{region "07 - Consume Start and Abort without restarting"}
FSteps[7].ExpectedState := E_State.Completed;
FSteps[7].ExpectedResult := E_Result.Passed;
FSteps[7].ExpectedReady := FALSE;
FSteps[7].ExpectedPassedCount := 2;
FSteps[7].ExpectedFailedCount := 0;
FSteps[7].CheckFinalization := TRUE;
FSteps[7].ExpectedFinalizationCount := 1;
FSteps[7].ExpectedCompletionCount := 1;
FSteps[7].ExpectedFinalResult := E_Result.Passed;
FSteps[7].ExpectRuntimeHeld := TRUE;
FSteps[7].RequestStart := TRUE;
FSteps[7].RequestAbort := TRUE;
FSteps[7].ExpectedHookCount := 1;
FSteps[7].ExpectedHooks[1].Hook := E_LifecycleHook.Aggregate;
FSteps[7].ExpectedHooks[1].State := E_State.Completed;
FSteps[7].ExpectedHooks[1].Enabled := TRUE;
{endregion}

{region "08 - Remain quiet after rejected terminal requests"}
FSteps[8].ExpectedState := E_State.Completed;
FSteps[8].ExpectedResult := E_Result.Passed;
FSteps[8].ExpectedReady := FALSE;
FSteps[8].ExpectedPassedCount := 2;
FSteps[8].ExpectedFailedCount := 0;
FSteps[8].CheckFinalization := TRUE;
FSteps[8].ExpectedFinalizationCount := 1;
FSteps[8].ExpectedCompletionCount := 1;
FSteps[8].ExpectedFinalResult := E_Result.Passed;
FSteps[8].ExpectRuntimeHeld := TRUE;
FSteps[8].ExpectQuietCall := TRUE;
FSteps[8].ExpectedHookCount := 1;
FSteps[8].ExpectedHooks[1].Hook := E_LifecycleHook.Aggregate;
FSteps[8].ExpectedHooks[1].State := E_State.Completed;
FSteps[8].ExpectedHooks[1].Enabled := TRUE;
{endregion}

{region "09 - Reset clears the first result and competing requests"}
FSteps[9].ExpectedState := E_State.Idle;
FSteps[9].ExpectedResult := E_Result.NotEvaluated;
FSteps[9].ExpectedReady := TRUE;
FSteps[9].ExpectedPassedCount := 0;
FSteps[9].ExpectedFailedCount := 0;
FSteps[9].CheckFinalization := TRUE;
FSteps[9].ExpectedFinalizationCount := 1;
FSteps[9].ExpectedCompletionCount := 1;
FSteps[9].ExpectedFinalResult := E_Result.Passed;
FSteps[9].RequestReset := TRUE;
FSteps[9].RequestStart := TRUE;
FSteps[9].RequestAbort := TRUE;
FSteps[9].ExpectRuntimeCleared := TRUE;
FSteps[9].ExpectedHookCount := 6;
FSteps[9].ExpectedHooks[1].Hook := E_LifecycleHook.Reset;
FSteps[9].ExpectedHooks[1].State := E_State.Reset;
FSteps[9].ExpectedHooks[1].Enabled := TRUE;
FSteps[9].ExpectedHooks[2].Hook := E_LifecycleHook.Abort;
FSteps[9].ExpectedHooks[2].State := E_State.Idle;
FSteps[9].ExpectedHooks[2].Enabled := FALSE;
FSteps[9].ExpectedHooks[3].Hook := E_LifecycleHook.Preparations;
FSteps[9].ExpectedHooks[3].State := E_State.Idle;
FSteps[9].ExpectedHooks[3].Enabled := FALSE;
FSteps[9].ExpectedHooks[4].Hook := E_LifecycleHook.Tests;
FSteps[9].ExpectedHooks[4].State := E_State.Idle;
FSteps[9].ExpectedHooks[4].Enabled := FALSE;
FSteps[9].ExpectedHooks[5].Hook := E_LifecycleHook.Assertions;
FSteps[9].ExpectedHooks[5].State := E_State.Idle;
FSteps[9].ExpectedHooks[5].Enabled := FALSE;
FSteps[9].ExpectedHooks[6].Hook := E_LifecycleHook.Aggregate;
FSteps[9].ExpectedHooks[6].State := E_State.Idle;
FSteps[9].ExpectedHooks[6].Enabled := TRUE;
{endregion}

{region "10 - Do not retain a Start from the Reset call"}
FSteps[10].ExpectedState := E_State.Idle;
FSteps[10].ExpectedResult := E_Result.NotEvaluated;
FSteps[10].ExpectedReady := TRUE;
FSteps[10].ExpectedPassedCount := 0;
FSteps[10].ExpectedFailedCount := 0;
FSteps[10].CheckFinalization := TRUE;
FSteps[10].ExpectedFinalizationCount := 1;
FSteps[10].ExpectedCompletionCount := 1;
FSteps[10].ExpectedFinalResult := E_Result.Passed;
FSteps[10].ExpectRuntimeCleared := TRUE;
FSteps[10].ExpectQuietCall := TRUE;
FSteps[10].ExpectedHookCount := 5;
FSteps[10].ExpectedHooks[1].Hook := E_LifecycleHook.Abort;
FSteps[10].ExpectedHooks[1].State := E_State.Idle;
FSteps[10].ExpectedHooks[1].Enabled := FALSE;
FSteps[10].ExpectedHooks[2].Hook := E_LifecycleHook.Preparations;
FSteps[10].ExpectedHooks[2].State := E_State.Idle;
FSteps[10].ExpectedHooks[2].Enabled := FALSE;
FSteps[10].ExpectedHooks[3].Hook := E_LifecycleHook.Tests;
FSteps[10].ExpectedHooks[3].State := E_State.Idle;
FSteps[10].ExpectedHooks[3].Enabled := FALSE;
FSteps[10].ExpectedHooks[4].Hook := E_LifecycleHook.Assertions;
FSteps[10].ExpectedHooks[4].State := E_State.Idle;
FSteps[10].ExpectedHooks[4].Enabled := FALSE;
FSteps[10].ExpectedHooks[5].Hook := E_LifecycleHook.Aggregate;
FSteps[10].ExpectedHooks[5].State := E_State.Idle;
FSteps[10].ExpectedHooks[5].Enabled := TRUE;
{endregion}

{region "11 - Start a fresh second execution"}
FSteps[11].ExpectedState := E_State.Starting;
FSteps[11].ExpectedResult := E_Result.NotEvaluated;
FSteps[11].ExpectedReady := FALSE;
FSteps[11].ExpectedPassedCount := 0;
FSteps[11].ExpectedFailedCount := 0;
FSteps[11].CheckFinalization := TRUE;
FSteps[11].ExpectedFinalizationCount := 1;
FSteps[11].ExpectedCompletionCount := 1;
FSteps[11].ExpectedFinalResult := E_Result.Passed;
FSteps[11].RequestStart := TRUE;
FSteps[11].ExpectedHookCount := 5;
FSteps[11].ExpectedHooks[1].Hook := E_LifecycleHook.Abort;
FSteps[11].ExpectedHooks[1].State := E_State.Starting;
FSteps[11].ExpectedHooks[1].Enabled := FALSE;
FSteps[11].ExpectedHooks[2].Hook := E_LifecycleHook.Preparations;
FSteps[11].ExpectedHooks[2].State := E_State.Starting;
FSteps[11].ExpectedHooks[2].Enabled := FALSE;
FSteps[11].ExpectedHooks[3].Hook := E_LifecycleHook.Tests;
FSteps[11].ExpectedHooks[3].State := E_State.Starting;
FSteps[11].ExpectedHooks[3].Enabled := FALSE;
FSteps[11].ExpectedHooks[4].Hook := E_LifecycleHook.Assertions;
FSteps[11].ExpectedHooks[4].State := E_State.Starting;
FSteps[11].ExpectedHooks[4].Enabled := FALSE;
FSteps[11].ExpectedHooks[5].Hook := E_LifecycleHook.Aggregate;
FSteps[11].ExpectedHooks[5].State := E_State.Starting;
FSteps[11].ExpectedHooks[5].Enabled := TRUE;
{endregion}

{region "12 - Both Assertions pass after Reset"}
FSteps[12].ExpectedState := E_State.Running;
FSteps[12].ExpectedResult := E_Result.NotEvaluated;
FSteps[12].ExpectedReady := FALSE;
FSteps[12].ExpectedPassedCount := 2;
FSteps[12].ExpectedFailedCount := 0;
FSteps[12].CheckFinalization := TRUE;
FSteps[12].ExpectedFinalizationCount := 1;
FSteps[12].ExpectedCompletionCount := 1;
FSteps[12].ExpectedFinalResult := E_Result.Passed;
FSteps[12].ExpectedHookCount := 5;
FSteps[12].ExpectedHooks[1].Hook := E_LifecycleHook.Abort;
FSteps[12].ExpectedHooks[1].State := E_State.Running;
FSteps[12].ExpectedHooks[1].Enabled := FALSE;
FSteps[12].ExpectedHooks[2].Hook := E_LifecycleHook.Preparations;
FSteps[12].ExpectedHooks[2].State := E_State.Running;
FSteps[12].ExpectedHooks[2].Enabled := FALSE;
FSteps[12].ExpectedHooks[3].Hook := E_LifecycleHook.Tests;
FSteps[12].ExpectedHooks[3].State := E_State.Running;
FSteps[12].ExpectedHooks[3].Enabled := TRUE;
FSteps[12].ExpectedHooks[4].Hook := E_LifecycleHook.Assertions;
FSteps[12].ExpectedHooks[4].State := E_State.Running;
FSteps[12].ExpectedHooks[4].Enabled := TRUE;
FSteps[12].ExpectedHooks[5].Hook := E_LifecycleHook.Aggregate;
FSteps[12].ExpectedHooks[5].State := E_State.Running;
FSteps[12].ExpectedHooks[5].Enabled := TRUE;
{endregion}

{region "13 - Publish a new successful finalization"}
FSteps[13].ExpectedState := E_State.Completing;
FSteps[13].ExpectedResult := E_Result.Passed;
FSteps[13].ExpectedReady := FALSE;
FSteps[13].ExpectedPassedCount := 2;
FSteps[13].ExpectedFailedCount := 0;
FSteps[13].FinishTests := TRUE;
FSteps[13].CheckFinalization := TRUE;
FSteps[13].ExpectedFinalizationCount := 2;
FSteps[13].ExpectedCompletionCount := 1;
FSteps[13].ExpectedFinalResult := E_Result.Passed;
FSteps[13].ExpectedHookCount := 5;
FSteps[13].ExpectedHooks[1].Hook := E_LifecycleHook.Abort;
FSteps[13].ExpectedHooks[1].State := E_State.Running;
FSteps[13].ExpectedHooks[1].Enabled := FALSE;
FSteps[13].ExpectedHooks[2].Hook := E_LifecycleHook.Preparations;
FSteps[13].ExpectedHooks[2].State := E_State.Running;
FSteps[13].ExpectedHooks[2].Enabled := FALSE;
FSteps[13].ExpectedHooks[3].Hook := E_LifecycleHook.Tests;
FSteps[13].ExpectedHooks[3].State := E_State.Running;
FSteps[13].ExpectedHooks[3].Enabled := TRUE;
FSteps[13].ExpectedHooks[4].Hook := E_LifecycleHook.Assertions;
FSteps[13].ExpectedHooks[4].State := E_State.Completing;
FSteps[13].ExpectedHooks[4].Enabled := FALSE;
FSteps[13].ExpectedHooks[5].Hook := E_LifecycleHook.Aggregate;
FSteps[13].ExpectedHooks[5].State := E_State.Completing;
FSteps[13].ExpectedHooks[5].Enabled := TRUE;
{endregion}

{region "14 - Complete the second execution"}
FSteps[14].ExpectedState := E_State.Completed;
FSteps[14].ExpectedResult := E_Result.Passed;
FSteps[14].ExpectedReady := FALSE;
FSteps[14].ExpectedPassedCount := 2;
FSteps[14].ExpectedFailedCount := 0;
FSteps[14].ExpectRuntimeHeld := TRUE;
FSteps[14].CheckFinalization := TRUE;
FSteps[14].ExpectedFinalizationCount := 2;
FSteps[14].ExpectedCompletionCount := 2;
FSteps[14].ExpectedFinalResult := E_Result.Passed;
FSteps[14].ExpectedHookCount := 1;
FSteps[14].ExpectedHooks[1].Hook := E_LifecycleHook.Aggregate;
FSteps[14].ExpectedHooks[1].State := E_State.Completed;
FSteps[14].ExpectedHooks[1].Enabled := TRUE;
{endregion}

{region "15 - Do not repeat second-run finalization"}
FSteps[15].ExpectedState := E_State.Completed;
FSteps[15].ExpectedResult := E_Result.Passed;
FSteps[15].ExpectedReady := FALSE;
FSteps[15].ExpectedPassedCount := 2;
FSteps[15].ExpectedFailedCount := 0;
FSteps[15].ExpectQuietCall := TRUE;
FSteps[15].ExpectRuntimeHeld := TRUE;
FSteps[15].CheckFinalization := TRUE;
FSteps[15].ExpectedFinalizationCount := 2;
FSteps[15].ExpectedCompletionCount := 2;
FSteps[15].ExpectedFinalResult := E_Result.Passed;
FSteps[15].ExpectedHookCount := 1;
FSteps[15].ExpectedHooks[1].Hook := E_LifecycleHook.Aggregate;
FSteps[15].ExpectedHooks[1].State := E_State.Completed;
FSteps[15].ExpectedHooks[1].Enabled := TRUE;
{endregion}
END_METHOD

END_FUNCTION_BLOCK

// ---- SelfTests/TestCases/TestSuite_TestCaseLifecycle/Test_LifecycleRepeatAfterFailed.TcPOU
{region 'Documentation'}
(*!
<summary>Checks stable Failed completion, one-shot finalization and a fresh successful run after Reset.</summary>
*)
{endregion}
FUNCTION_BLOCK Test_LifecycleRepeatAfterFailed EXTENDS TestCaseLifecycleTestBase

SUPER^();

{region 'Documentation'}
(*!
<summary>Defines two independent run outcomes and cumulative event expectations across Reset.</summary>
*)
{endregion}
METHOD PROTECTED ConfigureScenario
FSubjectPreparationCount := 0;
FSubjectTestCount := 1;
FStepCount := 15;

{region "01 - Reset establishes the initial Idle state"}
FSteps[1].ExpectedState := E_State.Idle;
FSteps[1].ExpectedResult := E_Result.NotEvaluated;
FSteps[1].ExpectedReady := TRUE;
FSteps[1].ExpectedPassedCount := 0;
FSteps[1].ExpectedFailedCount := 0;
FSteps[1].RequestReset := TRUE;
FSteps[1].ExpectRuntimeCleared := TRUE;
FSteps[1].CheckFinalization := TRUE;
FSteps[1].ExpectedFinalizationCount := 0;
FSteps[1].ExpectedCompletionCount := 0;
FSteps[1].ExpectedFinalResult := E_Result.Failed;
FSteps[1].ExpectedHookCount := 6;
FSteps[1].ExpectedHooks[1].Hook := E_LifecycleHook.Reset;
FSteps[1].ExpectedHooks[1].State := E_State.Reset;
FSteps[1].ExpectedHooks[1].Enabled := TRUE;
FSteps[1].ExpectedHooks[2].Hook := E_LifecycleHook.Abort;
FSteps[1].ExpectedHooks[2].State := E_State.Idle;
FSteps[1].ExpectedHooks[2].Enabled := FALSE;
FSteps[1].ExpectedHooks[3].Hook := E_LifecycleHook.Preparations;
FSteps[1].ExpectedHooks[3].State := E_State.Idle;
FSteps[1].ExpectedHooks[3].Enabled := FALSE;
FSteps[1].ExpectedHooks[4].Hook := E_LifecycleHook.Tests;
FSteps[1].ExpectedHooks[4].State := E_State.Idle;
FSteps[1].ExpectedHooks[4].Enabled := FALSE;
FSteps[1].ExpectedHooks[5].Hook := E_LifecycleHook.Assertions;
FSteps[1].ExpectedHooks[5].State := E_State.Idle;
FSteps[1].ExpectedHooks[5].Enabled := FALSE;
FSteps[1].ExpectedHooks[6].Hook := E_LifecycleHook.Aggregate;
FSteps[1].ExpectedHooks[6].State := E_State.Idle;
FSteps[1].ExpectedHooks[6].Enabled := TRUE;
{endregion}

{region "02 - Start the first execution"}
FSteps[2].ExpectedState := E_State.Starting;
FSteps[2].ExpectedResult := E_Result.NotEvaluated;
FSteps[2].ExpectedReady := FALSE;
FSteps[2].ExpectedPassedCount := 0;
FSteps[2].ExpectedFailedCount := 0;
FSteps[2].RequestStart := TRUE;
FSteps[2].CheckFinalization := TRUE;
FSteps[2].ExpectedFinalizationCount := 0;
FSteps[2].ExpectedCompletionCount := 0;
FSteps[2].ExpectedFinalResult := E_Result.Failed;
FSteps[2].ExpectedHookCount := 5;
FSteps[2].ExpectedHooks[1].Hook := E_LifecycleHook.Abort;
FSteps[2].ExpectedHooks[1].State := E_State.Starting;
FSteps[2].ExpectedHooks[1].Enabled := FALSE;
FSteps[2].ExpectedHooks[2].Hook := E_LifecycleHook.Preparations;
FSteps[2].ExpectedHooks[2].State := E_State.Starting;
FSteps[2].ExpectedHooks[2].Enabled := FALSE;
FSteps[2].ExpectedHooks[3].Hook := E_LifecycleHook.Tests;
FSteps[2].ExpectedHooks[3].State := E_State.Starting;
FSteps[2].ExpectedHooks[3].Enabled := FALSE;
FSteps[2].ExpectedHooks[4].Hook := E_LifecycleHook.Assertions;
FSteps[2].ExpectedHooks[4].State := E_State.Starting;
FSteps[2].ExpectedHooks[4].Enabled := FALSE;
FSteps[2].ExpectedHooks[5].Hook := E_LifecycleHook.Aggregate;
FSteps[2].ExpectedHooks[5].State := E_State.Starting;
FSteps[2].ExpectedHooks[5].Enabled := TRUE;
{endregion}

{region "03 - Evaluate both child Assertions"}
FSteps[3].ExpectedState := E_State.Running;
FSteps[3].ExpectedResult := E_Result.NotEvaluated;
FSteps[3].ExpectedReady := FALSE;
FSteps[3].ExpectedPassedCount := 1;
FSteps[3].ExpectedFailedCount := 1;
FSteps[3].AssertionCondition := FALSE;
FSteps[3].CheckFinalization := TRUE;
FSteps[3].ExpectedFinalizationCount := 0;
FSteps[3].ExpectedCompletionCount := 0;
FSteps[3].ExpectedFinalResult := E_Result.Failed;
FSteps[3].ExpectedHookCount := 5;
FSteps[3].ExpectedHooks[1].Hook := E_LifecycleHook.Abort;
FSteps[3].ExpectedHooks[1].State := E_State.Running;
FSteps[3].ExpectedHooks[1].Enabled := FALSE;
FSteps[3].ExpectedHooks[2].Hook := E_LifecycleHook.Preparations;
FSteps[3].ExpectedHooks[2].State := E_State.Running;
FSteps[3].ExpectedHooks[2].Enabled := FALSE;
FSteps[3].ExpectedHooks[3].Hook := E_LifecycleHook.Tests;
FSteps[3].ExpectedHooks[3].State := E_State.Running;
FSteps[3].ExpectedHooks[3].Enabled := TRUE;
FSteps[3].ExpectedHooks[4].Hook := E_LifecycleHook.Assertions;
FSteps[3].ExpectedHooks[4].State := E_State.Running;
FSteps[3].ExpectedHooks[4].Enabled := TRUE;
FSteps[3].ExpectedHooks[5].Hook := E_LifecycleHook.Aggregate;
FSteps[3].ExpectedHooks[5].State := E_State.Running;
FSteps[3].ExpectedHooks[5].Enabled := TRUE;
{endregion}

{region "04 - Finalize the first result"}
FSteps[4].ExpectedState := E_State.Completing;
FSteps[4].ExpectedResult := E_Result.Failed;
FSteps[4].ExpectedReady := FALSE;
FSteps[4].ExpectedPassedCount := 1;
FSteps[4].ExpectedFailedCount := 1;
FSteps[4].FinishTests := TRUE;
FSteps[4].CheckFinalization := TRUE;
FSteps[4].ExpectedFinalizationCount := 1;
FSteps[4].ExpectedCompletionCount := 0;
FSteps[4].ExpectedFinalResult := E_Result.Failed;
FSteps[4].ExpectedHookCount := 5;
FSteps[4].ExpectedHooks[1].Hook := E_LifecycleHook.Abort;
FSteps[4].ExpectedHooks[1].State := E_State.Running;
FSteps[4].ExpectedHooks[1].Enabled := FALSE;
FSteps[4].ExpectedHooks[2].Hook := E_LifecycleHook.Preparations;
FSteps[4].ExpectedHooks[2].State := E_State.Running;
FSteps[4].ExpectedHooks[2].Enabled := FALSE;
FSteps[4].ExpectedHooks[3].Hook := E_LifecycleHook.Tests;
FSteps[4].ExpectedHooks[3].State := E_State.Running;
FSteps[4].ExpectedHooks[3].Enabled := TRUE;
FSteps[4].ExpectedHooks[4].Hook := E_LifecycleHook.Assertions;
FSteps[4].ExpectedHooks[4].State := E_State.Completing;
FSteps[4].ExpectedHooks[4].Enabled := FALSE;
FSteps[4].ExpectedHooks[5].Hook := E_LifecycleHook.Aggregate;
FSteps[4].ExpectedHooks[5].State := E_State.Completing;
FSteps[4].ExpectedHooks[5].Enabled := TRUE;
{endregion}

{region "05 - Observe the final Completed transition"}
FSteps[5].ExpectedState := E_State.Completed;
FSteps[5].ExpectedResult := E_Result.Failed;
FSteps[5].ExpectedReady := FALSE;
FSteps[5].ExpectedPassedCount := 1;
FSteps[5].ExpectedFailedCount := 1;
FSteps[5].CheckFinalization := TRUE;
FSteps[5].ExpectedFinalizationCount := 1;
FSteps[5].ExpectedCompletionCount := 1;
FSteps[5].ExpectedFinalResult := E_Result.Failed;
FSteps[5].ExpectRuntimeHeld := TRUE;
FSteps[5].ExpectedHookCount := 1;
FSteps[5].ExpectedHooks[1].Hook := E_LifecycleHook.Aggregate;
FSteps[5].ExpectedHooks[1].State := E_State.Completed;
FSteps[5].ExpectedHooks[1].Enabled := TRUE;
{endregion}

{region "06 - Ignore processing inputs while Completed"}
FSteps[6].ExpectedState := E_State.Completed;
FSteps[6].ExpectedResult := E_Result.Failed;
FSteps[6].ExpectedReady := FALSE;
FSteps[6].ExpectedPassedCount := 1;
FSteps[6].ExpectedFailedCount := 1;
FSteps[6].CheckFinalization := TRUE;
FSteps[6].ExpectedFinalizationCount := 1;
FSteps[6].ExpectedCompletionCount := 1;
FSteps[6].ExpectedFinalResult := E_Result.Failed;
FSteps[6].ExpectRuntimeHeld := TRUE;
FSteps[6].ExpectQuietCall := TRUE;
FSteps[6].Ready := FALSE;
FSteps[6].ResetError := TRUE;
FSteps[6].AbortError := TRUE;
FSteps[6].TestError := TRUE;
FSteps[6].PreparationError := TRUE;
FSteps[6].AdvancePreparation := TRUE;
FSteps[6].FinishPreparations := TRUE;
FSteps[6].AdvanceTest := TRUE;
FSteps[6].FinishTests := TRUE;
FSteps[6].AssertionCondition := FALSE;
FSteps[6].ExpectedHookCount := 1;
FSteps[6].ExpectedHooks[1].Hook := E_LifecycleHook.Aggregate;
FSteps[6].ExpectedHooks[1].State := E_State.Completed;
FSteps[6].ExpectedHooks[1].Enabled := TRUE;
{endregion}

{region "07 - Consume Start and Abort without restarting"}
FSteps[7].ExpectedState := E_State.Completed;
FSteps[7].ExpectedResult := E_Result.Failed;
FSteps[7].ExpectedReady := FALSE;
FSteps[7].ExpectedPassedCount := 1;
FSteps[7].ExpectedFailedCount := 1;
FSteps[7].CheckFinalization := TRUE;
FSteps[7].ExpectedFinalizationCount := 1;
FSteps[7].ExpectedCompletionCount := 1;
FSteps[7].ExpectedFinalResult := E_Result.Failed;
FSteps[7].ExpectRuntimeHeld := TRUE;
FSteps[7].RequestStart := TRUE;
FSteps[7].RequestAbort := TRUE;
FSteps[7].ExpectedHookCount := 1;
FSteps[7].ExpectedHooks[1].Hook := E_LifecycleHook.Aggregate;
FSteps[7].ExpectedHooks[1].State := E_State.Completed;
FSteps[7].ExpectedHooks[1].Enabled := TRUE;
{endregion}

{region "08 - Remain quiet after rejected terminal requests"}
FSteps[8].ExpectedState := E_State.Completed;
FSteps[8].ExpectedResult := E_Result.Failed;
FSteps[8].ExpectedReady := FALSE;
FSteps[8].ExpectedPassedCount := 1;
FSteps[8].ExpectedFailedCount := 1;
FSteps[8].CheckFinalization := TRUE;
FSteps[8].ExpectedFinalizationCount := 1;
FSteps[8].ExpectedCompletionCount := 1;
FSteps[8].ExpectedFinalResult := E_Result.Failed;
FSteps[8].ExpectRuntimeHeld := TRUE;
FSteps[8].ExpectQuietCall := TRUE;
FSteps[8].ExpectedHookCount := 1;
FSteps[8].ExpectedHooks[1].Hook := E_LifecycleHook.Aggregate;
FSteps[8].ExpectedHooks[1].State := E_State.Completed;
FSteps[8].ExpectedHooks[1].Enabled := TRUE;
{endregion}

{region "09 - Reset clears the first result and competing requests"}
FSteps[9].ExpectedState := E_State.Idle;
FSteps[9].ExpectedResult := E_Result.NotEvaluated;
FSteps[9].ExpectedReady := TRUE;
FSteps[9].ExpectedPassedCount := 0;
FSteps[9].ExpectedFailedCount := 0;
FSteps[9].CheckFinalization := TRUE;
FSteps[9].ExpectedFinalizationCount := 1;
FSteps[9].ExpectedCompletionCount := 1;
FSteps[9].ExpectedFinalResult := E_Result.Failed;
FSteps[9].RequestReset := TRUE;
FSteps[9].RequestStart := TRUE;
FSteps[9].RequestAbort := TRUE;
FSteps[9].ExpectRuntimeCleared := TRUE;
FSteps[9].ExpectedHookCount := 6;
FSteps[9].ExpectedHooks[1].Hook := E_LifecycleHook.Reset;
FSteps[9].ExpectedHooks[1].State := E_State.Reset;
FSteps[9].ExpectedHooks[1].Enabled := TRUE;
FSteps[9].ExpectedHooks[2].Hook := E_LifecycleHook.Abort;
FSteps[9].ExpectedHooks[2].State := E_State.Idle;
FSteps[9].ExpectedHooks[2].Enabled := FALSE;
FSteps[9].ExpectedHooks[3].Hook := E_LifecycleHook.Preparations;
FSteps[9].ExpectedHooks[3].State := E_State.Idle;
FSteps[9].ExpectedHooks[3].Enabled := FALSE;
FSteps[9].ExpectedHooks[4].Hook := E_LifecycleHook.Tests;
FSteps[9].ExpectedHooks[4].State := E_State.Idle;
FSteps[9].ExpectedHooks[4].Enabled := FALSE;
FSteps[9].ExpectedHooks[5].Hook := E_LifecycleHook.Assertions;
FSteps[9].ExpectedHooks[5].State := E_State.Idle;
FSteps[9].ExpectedHooks[5].Enabled := FALSE;
FSteps[9].ExpectedHooks[6].Hook := E_LifecycleHook.Aggregate;
FSteps[9].ExpectedHooks[6].State := E_State.Idle;
FSteps[9].ExpectedHooks[6].Enabled := TRUE;
{endregion}

{region "10 - Do not retain a Start from the Reset call"}
FSteps[10].ExpectedState := E_State.Idle;
FSteps[10].ExpectedResult := E_Result.NotEvaluated;
FSteps[10].ExpectedReady := TRUE;
FSteps[10].ExpectedPassedCount := 0;
FSteps[10].ExpectedFailedCount := 0;
FSteps[10].CheckFinalization := TRUE;
FSteps[10].ExpectedFinalizationCount := 1;
FSteps[10].ExpectedCompletionCount := 1;
FSteps[10].ExpectedFinalResult := E_Result.Failed;
FSteps[10].ExpectRuntimeCleared := TRUE;
FSteps[10].ExpectQuietCall := TRUE;
FSteps[10].ExpectedHookCount := 5;
FSteps[10].ExpectedHooks[1].Hook := E_LifecycleHook.Abort;
FSteps[10].ExpectedHooks[1].State := E_State.Idle;
FSteps[10].ExpectedHooks[1].Enabled := FALSE;
FSteps[10].ExpectedHooks[2].Hook := E_LifecycleHook.Preparations;
FSteps[10].ExpectedHooks[2].State := E_State.Idle;
FSteps[10].ExpectedHooks[2].Enabled := FALSE;
FSteps[10].ExpectedHooks[3].Hook := E_LifecycleHook.Tests;
FSteps[10].ExpectedHooks[3].State := E_State.Idle;
FSteps[10].ExpectedHooks[3].Enabled := FALSE;
FSteps[10].ExpectedHooks[4].Hook := E_LifecycleHook.Assertions;
FSteps[10].ExpectedHooks[4].State := E_State.Idle;
FSteps[10].ExpectedHooks[4].Enabled := FALSE;
FSteps[10].ExpectedHooks[5].Hook := E_LifecycleHook.Aggregate;
FSteps[10].ExpectedHooks[5].State := E_State.Idle;
FSteps[10].ExpectedHooks[5].Enabled := TRUE;
{endregion}

{region "11 - Start a fresh second execution"}
FSteps[11].ExpectedState := E_State.Starting;
FSteps[11].ExpectedResult := E_Result.NotEvaluated;
FSteps[11].ExpectedReady := FALSE;
FSteps[11].ExpectedPassedCount := 0;
FSteps[11].ExpectedFailedCount := 0;
FSteps[11].CheckFinalization := TRUE;
FSteps[11].ExpectedFinalizationCount := 1;
FSteps[11].ExpectedCompletionCount := 1;
FSteps[11].ExpectedFinalResult := E_Result.Failed;
FSteps[11].RequestStart := TRUE;
FSteps[11].ExpectedHookCount := 5;
FSteps[11].ExpectedHooks[1].Hook := E_LifecycleHook.Abort;
FSteps[11].ExpectedHooks[1].State := E_State.Starting;
FSteps[11].ExpectedHooks[1].Enabled := FALSE;
FSteps[11].ExpectedHooks[2].Hook := E_LifecycleHook.Preparations;
FSteps[11].ExpectedHooks[2].State := E_State.Starting;
FSteps[11].ExpectedHooks[2].Enabled := FALSE;
FSteps[11].ExpectedHooks[3].Hook := E_LifecycleHook.Tests;
FSteps[11].ExpectedHooks[3].State := E_State.Starting;
FSteps[11].ExpectedHooks[3].Enabled := FALSE;
FSteps[11].ExpectedHooks[4].Hook := E_LifecycleHook.Assertions;
FSteps[11].ExpectedHooks[4].State := E_State.Starting;
FSteps[11].ExpectedHooks[4].Enabled := FALSE;
FSteps[11].ExpectedHooks[5].Hook := E_LifecycleHook.Aggregate;
FSteps[11].ExpectedHooks[5].State := E_State.Starting;
FSteps[11].ExpectedHooks[5].Enabled := TRUE;
{endregion}

{region "12 - Both Assertions pass after Reset"}
FSteps[12].ExpectedState := E_State.Running;
FSteps[12].ExpectedResult := E_Result.NotEvaluated;
FSteps[12].ExpectedReady := FALSE;
FSteps[12].ExpectedPassedCount := 2;
FSteps[12].ExpectedFailedCount := 0;
FSteps[12].CheckFinalization := TRUE;
FSteps[12].ExpectedFinalizationCount := 1;
FSteps[12].ExpectedCompletionCount := 1;
FSteps[12].ExpectedFinalResult := E_Result.Failed;
FSteps[12].ExpectedHookCount := 5;
FSteps[12].ExpectedHooks[1].Hook := E_LifecycleHook.Abort;
FSteps[12].ExpectedHooks[1].State := E_State.Running;
FSteps[12].ExpectedHooks[1].Enabled := FALSE;
FSteps[12].ExpectedHooks[2].Hook := E_LifecycleHook.Preparations;
FSteps[12].ExpectedHooks[2].State := E_State.Running;
FSteps[12].ExpectedHooks[2].Enabled := FALSE;
FSteps[12].ExpectedHooks[3].Hook := E_LifecycleHook.Tests;
FSteps[12].ExpectedHooks[3].State := E_State.Running;
FSteps[12].ExpectedHooks[3].Enabled := TRUE;
FSteps[12].ExpectedHooks[4].Hook := E_LifecycleHook.Assertions;
FSteps[12].ExpectedHooks[4].State := E_State.Running;
FSteps[12].ExpectedHooks[4].Enabled := TRUE;
FSteps[12].ExpectedHooks[5].Hook := E_LifecycleHook.Aggregate;
FSteps[12].ExpectedHooks[5].State := E_State.Running;
FSteps[12].ExpectedHooks[5].Enabled := TRUE;
{endregion}

{region "13 - Publish a new successful finalization"}
FSteps[13].ExpectedState := E_State.Completing;
FSteps[13].ExpectedResult := E_Result.Passed;
FSteps[13].ExpectedReady := FALSE;
FSteps[13].ExpectedPassedCount := 2;
FSteps[13].ExpectedFailedCount := 0;
FSteps[13].FinishTests := TRUE;
FSteps[13].CheckFinalization := TRUE;
FSteps[13].ExpectedFinalizationCount := 2;
FSteps[13].ExpectedCompletionCount := 1;
FSteps[13].ExpectedFinalResult := E_Result.Passed;
FSteps[13].ExpectedHookCount := 5;
FSteps[13].ExpectedHooks[1].Hook := E_LifecycleHook.Abort;
FSteps[13].ExpectedHooks[1].State := E_State.Running;
FSteps[13].ExpectedHooks[1].Enabled := FALSE;
FSteps[13].ExpectedHooks[2].Hook := E_LifecycleHook.Preparations;
FSteps[13].ExpectedHooks[2].State := E_State.Running;
FSteps[13].ExpectedHooks[2].Enabled := FALSE;
FSteps[13].ExpectedHooks[3].Hook := E_LifecycleHook.Tests;
FSteps[13].ExpectedHooks[3].State := E_State.Running;
FSteps[13].ExpectedHooks[3].Enabled := TRUE;
FSteps[13].ExpectedHooks[4].Hook := E_LifecycleHook.Assertions;
FSteps[13].ExpectedHooks[4].State := E_State.Completing;
FSteps[13].ExpectedHooks[4].Enabled := FALSE;
FSteps[13].ExpectedHooks[5].Hook := E_LifecycleHook.Aggregate;
FSteps[13].ExpectedHooks[5].State := E_State.Completing;
FSteps[13].ExpectedHooks[5].Enabled := TRUE;
{endregion}

{region "14 - Complete the second execution"}
FSteps[14].ExpectedState := E_State.Completed;
FSteps[14].ExpectedResult := E_Result.Passed;
FSteps[14].ExpectedReady := FALSE;
FSteps[14].ExpectedPassedCount := 2;
FSteps[14].ExpectedFailedCount := 0;
FSteps[14].ExpectRuntimeHeld := TRUE;
FSteps[14].CheckFinalization := TRUE;
FSteps[14].ExpectedFinalizationCount := 2;
FSteps[14].ExpectedCompletionCount := 2;
FSteps[14].ExpectedFinalResult := E_Result.Passed;
FSteps[14].ExpectedHookCount := 1;
FSteps[14].ExpectedHooks[1].Hook := E_LifecycleHook.Aggregate;
FSteps[14].ExpectedHooks[1].State := E_State.Completed;
FSteps[14].ExpectedHooks[1].Enabled := TRUE;
{endregion}

{region "15 - Do not repeat second-run finalization"}
FSteps[15].ExpectedState := E_State.Completed;
FSteps[15].ExpectedResult := E_Result.Passed;
FSteps[15].ExpectedReady := FALSE;
FSteps[15].ExpectedPassedCount := 2;
FSteps[15].ExpectedFailedCount := 0;
FSteps[15].ExpectQuietCall := TRUE;
FSteps[15].ExpectRuntimeHeld := TRUE;
FSteps[15].CheckFinalization := TRUE;
FSteps[15].ExpectedFinalizationCount := 2;
FSteps[15].ExpectedCompletionCount := 2;
FSteps[15].ExpectedFinalResult := E_Result.Passed;
FSteps[15].ExpectedHookCount := 1;
FSteps[15].ExpectedHooks[1].Hook := E_LifecycleHook.Aggregate;
FSteps[15].ExpectedHooks[1].State := E_State.Completed;
FSteps[15].ExpectedHooks[1].Enabled := TRUE;
{endregion}
END_METHOD

END_FUNCTION_BLOCK

// ---- SelfTests/TestCases/TestSuite_TestCaseLifecycle/Test_LifecycleRepeatAfterError.TcPOU
{region 'Documentation'}
(*!
<summary>Checks stable Error completion, one-shot finalization and a fresh successful run after Reset.</summary>
*)
{endregion}
FUNCTION_BLOCK Test_LifecycleRepeatAfterError EXTENDS TestCaseLifecycleTestBase

SUPER^();

{region 'Documentation'}
(*!
<summary>Defines two independent run outcomes and cumulative event expectations across Reset.</summary>
*)
{endregion}
METHOD PROTECTED ConfigureScenario
FSubjectPreparationCount := 0;
FSubjectTestCount := 1;
FStepCount := 16;

{region "01 - Reset establishes the initial Idle state"}
FSteps[1].ExpectedState := E_State.Idle;
FSteps[1].ExpectedResult := E_Result.NotEvaluated;
FSteps[1].ExpectedReady := TRUE;
FSteps[1].ExpectedPassedCount := 0;
FSteps[1].ExpectedFailedCount := 0;
FSteps[1].RequestReset := TRUE;
FSteps[1].ExpectRuntimeCleared := TRUE;
FSteps[1].CheckFinalization := TRUE;
FSteps[1].ExpectedFinalizationCount := 0;
FSteps[1].ExpectedCompletionCount := 0;
FSteps[1].ExpectedFinalResult := E_Result.Error;
FSteps[1].ExpectedHookCount := 6;
FSteps[1].ExpectedHooks[1].Hook := E_LifecycleHook.Reset;
FSteps[1].ExpectedHooks[1].State := E_State.Reset;
FSteps[1].ExpectedHooks[1].Enabled := TRUE;
FSteps[1].ExpectedHooks[2].Hook := E_LifecycleHook.Abort;
FSteps[1].ExpectedHooks[2].State := E_State.Idle;
FSteps[1].ExpectedHooks[2].Enabled := FALSE;
FSteps[1].ExpectedHooks[3].Hook := E_LifecycleHook.Preparations;
FSteps[1].ExpectedHooks[3].State := E_State.Idle;
FSteps[1].ExpectedHooks[3].Enabled := FALSE;
FSteps[1].ExpectedHooks[4].Hook := E_LifecycleHook.Tests;
FSteps[1].ExpectedHooks[4].State := E_State.Idle;
FSteps[1].ExpectedHooks[4].Enabled := FALSE;
FSteps[1].ExpectedHooks[5].Hook := E_LifecycleHook.Assertions;
FSteps[1].ExpectedHooks[5].State := E_State.Idle;
FSteps[1].ExpectedHooks[5].Enabled := FALSE;
FSteps[1].ExpectedHooks[6].Hook := E_LifecycleHook.Aggregate;
FSteps[1].ExpectedHooks[6].State := E_State.Idle;
FSteps[1].ExpectedHooks[6].Enabled := TRUE;
{endregion}

{region "02 - Start the first execution"}
FSteps[2].ExpectedState := E_State.Starting;
FSteps[2].ExpectedResult := E_Result.NotEvaluated;
FSteps[2].ExpectedReady := FALSE;
FSteps[2].ExpectedPassedCount := 0;
FSteps[2].ExpectedFailedCount := 0;
FSteps[2].RequestStart := TRUE;
FSteps[2].CheckFinalization := TRUE;
FSteps[2].ExpectedFinalizationCount := 0;
FSteps[2].ExpectedCompletionCount := 0;
FSteps[2].ExpectedFinalResult := E_Result.Error;
FSteps[2].ExpectedHookCount := 5;
FSteps[2].ExpectedHooks[1].Hook := E_LifecycleHook.Abort;
FSteps[2].ExpectedHooks[1].State := E_State.Starting;
FSteps[2].ExpectedHooks[1].Enabled := FALSE;
FSteps[2].ExpectedHooks[2].Hook := E_LifecycleHook.Preparations;
FSteps[2].ExpectedHooks[2].State := E_State.Starting;
FSteps[2].ExpectedHooks[2].Enabled := FALSE;
FSteps[2].ExpectedHooks[3].Hook := E_LifecycleHook.Tests;
FSteps[2].ExpectedHooks[3].State := E_State.Starting;
FSteps[2].ExpectedHooks[3].Enabled := FALSE;
FSteps[2].ExpectedHooks[4].Hook := E_LifecycleHook.Assertions;
FSteps[2].ExpectedHooks[4].State := E_State.Starting;
FSteps[2].ExpectedHooks[4].Enabled := FALSE;
FSteps[2].ExpectedHooks[5].Hook := E_LifecycleHook.Aggregate;
FSteps[2].ExpectedHooks[5].State := E_State.Starting;
FSteps[2].ExpectedHooks[5].Enabled := TRUE;
{endregion}

{region "03 - Evaluate both child Assertions"}
FSteps[3].ExpectedState := E_State.Running;
FSteps[3].ExpectedResult := E_Result.NotEvaluated;
FSteps[3].ExpectedReady := FALSE;
FSteps[3].ExpectedPassedCount := 2;
FSteps[3].ExpectedFailedCount := 0;
FSteps[3].AssertionCondition := TRUE;
FSteps[3].CheckFinalization := TRUE;
FSteps[3].ExpectedFinalizationCount := 0;
FSteps[3].ExpectedCompletionCount := 0;
FSteps[3].ExpectedFinalResult := E_Result.Error;
FSteps[3].ExpectedHookCount := 5;
FSteps[3].ExpectedHooks[1].Hook := E_LifecycleHook.Abort;
FSteps[3].ExpectedHooks[1].State := E_State.Running;
FSteps[3].ExpectedHooks[1].Enabled := FALSE;
FSteps[3].ExpectedHooks[2].Hook := E_LifecycleHook.Preparations;
FSteps[3].ExpectedHooks[2].State := E_State.Running;
FSteps[3].ExpectedHooks[2].Enabled := FALSE;
FSteps[3].ExpectedHooks[3].Hook := E_LifecycleHook.Tests;
FSteps[3].ExpectedHooks[3].State := E_State.Running;
FSteps[3].ExpectedHooks[3].Enabled := TRUE;
FSteps[3].ExpectedHooks[4].Hook := E_LifecycleHook.Assertions;
FSteps[3].ExpectedHooks[4].State := E_State.Running;
FSteps[3].ExpectedHooks[4].Enabled := TRUE;
FSteps[3].ExpectedHooks[5].Hook := E_LifecycleHook.Aggregate;
FSteps[3].ExpectedHooks[5].State := E_State.Running;
FSteps[3].ExpectedHooks[5].Enabled := TRUE;
{endregion}

{region "04 - Escalate execution to Error"}
FSteps[4].ExpectedState := E_State.AbortingFromError;
FSteps[4].ExpectedResult := E_Result.Error;
FSteps[4].ExpectedReady := FALSE;
FSteps[4].ExpectedPassedCount := 2;
FSteps[4].ExpectedFailedCount := 0;
FSteps[4].TestError := TRUE;
FSteps[4].CheckFinalization := TRUE;
FSteps[4].ExpectedFinalizationCount := 0;
FSteps[4].ExpectedCompletionCount := 0;
FSteps[4].ExpectedFinalResult := E_Result.Error;
FSteps[4].ExpectedHookCount := 5;
FSteps[4].ExpectedHooks[1].Hook := E_LifecycleHook.Abort;
FSteps[4].ExpectedHooks[1].State := E_State.Running;
FSteps[4].ExpectedHooks[1].Enabled := FALSE;
FSteps[4].ExpectedHooks[2].Hook := E_LifecycleHook.Preparations;
FSteps[4].ExpectedHooks[2].State := E_State.Running;
FSteps[4].ExpectedHooks[2].Enabled := FALSE;
FSteps[4].ExpectedHooks[3].Hook := E_LifecycleHook.Tests;
FSteps[4].ExpectedHooks[3].State := E_State.Running;
FSteps[4].ExpectedHooks[3].Enabled := TRUE;
FSteps[4].ExpectedHooks[4].Hook := E_LifecycleHook.Assertions;
FSteps[4].ExpectedHooks[4].State := E_State.AbortingFromError;
FSteps[4].ExpectedHooks[4].Enabled := FALSE;
FSteps[4].ExpectedHooks[5].Hook := E_LifecycleHook.Aggregate;
FSteps[4].ExpectedHooks[5].State := E_State.AbortingFromError;
FSteps[4].ExpectedHooks[5].Enabled := TRUE;
{endregion}

{region "05 - Complete controlled Error cleanup"}
FSteps[5].ExpectedState := E_State.Completing;
FSteps[5].ExpectedResult := E_Result.Error;
FSteps[5].ExpectedReady := FALSE;
FSteps[5].ExpectedPassedCount := 2;
FSteps[5].ExpectedFailedCount := 0;
FSteps[5].CheckFinalization := TRUE;
FSteps[5].ExpectedFinalizationCount := 1;
FSteps[5].ExpectedCompletionCount := 0;
FSteps[5].ExpectedFinalResult := E_Result.Error;
FSteps[5].ExpectedHookCount := 5;
FSteps[5].ExpectedHooks[1].Hook := E_LifecycleHook.Abort;
FSteps[5].ExpectedHooks[1].State := E_State.AbortingFromError;
FSteps[5].ExpectedHooks[1].Enabled := TRUE;
FSteps[5].ExpectedHooks[2].Hook := E_LifecycleHook.Preparations;
FSteps[5].ExpectedHooks[2].State := E_State.Completing;
FSteps[5].ExpectedHooks[2].Enabled := FALSE;
FSteps[5].ExpectedHooks[3].Hook := E_LifecycleHook.Tests;
FSteps[5].ExpectedHooks[3].State := E_State.Completing;
FSteps[5].ExpectedHooks[3].Enabled := FALSE;
FSteps[5].ExpectedHooks[4].Hook := E_LifecycleHook.Assertions;
FSteps[5].ExpectedHooks[4].State := E_State.Completing;
FSteps[5].ExpectedHooks[4].Enabled := FALSE;
FSteps[5].ExpectedHooks[5].Hook := E_LifecycleHook.Aggregate;
FSteps[5].ExpectedHooks[5].State := E_State.Completing;
FSteps[5].ExpectedHooks[5].Enabled := TRUE;
{endregion}

{region "06 - Observe the final Completed transition"}
FSteps[6].ExpectedState := E_State.Completed;
FSteps[6].ExpectedResult := E_Result.Error;
FSteps[6].ExpectedReady := FALSE;
FSteps[6].ExpectedPassedCount := 2;
FSteps[6].ExpectedFailedCount := 0;
FSteps[6].CheckFinalization := TRUE;
FSteps[6].ExpectedFinalizationCount := 1;
FSteps[6].ExpectedCompletionCount := 1;
FSteps[6].ExpectedFinalResult := E_Result.Error;
FSteps[6].ExpectRuntimeHeld := TRUE;
FSteps[6].ExpectedHookCount := 1;
FSteps[6].ExpectedHooks[1].Hook := E_LifecycleHook.Aggregate;
FSteps[6].ExpectedHooks[1].State := E_State.Completed;
FSteps[6].ExpectedHooks[1].Enabled := TRUE;
{endregion}

{region "07 - Ignore processing inputs while Completed"}
FSteps[7].ExpectedState := E_State.Completed;
FSteps[7].ExpectedResult := E_Result.Error;
FSteps[7].ExpectedReady := FALSE;
FSteps[7].ExpectedPassedCount := 2;
FSteps[7].ExpectedFailedCount := 0;
FSteps[7].CheckFinalization := TRUE;
FSteps[7].ExpectedFinalizationCount := 1;
FSteps[7].ExpectedCompletionCount := 1;
FSteps[7].ExpectedFinalResult := E_Result.Error;
FSteps[7].ExpectRuntimeHeld := TRUE;
FSteps[7].ExpectQuietCall := TRUE;
FSteps[7].Ready := FALSE;
FSteps[7].ResetError := TRUE;
FSteps[7].AbortError := TRUE;
FSteps[7].TestError := TRUE;
FSteps[7].PreparationError := TRUE;
FSteps[7].AdvancePreparation := TRUE;
FSteps[7].FinishPreparations := TRUE;
FSteps[7].AdvanceTest := TRUE;
FSteps[7].FinishTests := TRUE;
FSteps[7].AssertionCondition := FALSE;
FSteps[7].ExpectedHookCount := 1;
FSteps[7].ExpectedHooks[1].Hook := E_LifecycleHook.Aggregate;
FSteps[7].ExpectedHooks[1].State := E_State.Completed;
FSteps[7].ExpectedHooks[1].Enabled := TRUE;
{endregion}

{region "08 - Consume Start and Abort without restarting"}
FSteps[8].ExpectedState := E_State.Completed;
FSteps[8].ExpectedResult := E_Result.Error;
FSteps[8].ExpectedReady := FALSE;
FSteps[8].ExpectedPassedCount := 2;
FSteps[8].ExpectedFailedCount := 0;
FSteps[8].CheckFinalization := TRUE;
FSteps[8].ExpectedFinalizationCount := 1;
FSteps[8].ExpectedCompletionCount := 1;
FSteps[8].ExpectedFinalResult := E_Result.Error;
FSteps[8].ExpectRuntimeHeld := TRUE;
FSteps[8].RequestStart := TRUE;
FSteps[8].RequestAbort := TRUE;
FSteps[8].ExpectedHookCount := 1;
FSteps[8].ExpectedHooks[1].Hook := E_LifecycleHook.Aggregate;
FSteps[8].ExpectedHooks[1].State := E_State.Completed;
FSteps[8].ExpectedHooks[1].Enabled := TRUE;
{endregion}

{region "09 - Remain quiet after rejected terminal requests"}
FSteps[9].ExpectedState := E_State.Completed;
FSteps[9].ExpectedResult := E_Result.Error;
FSteps[9].ExpectedReady := FALSE;
FSteps[9].ExpectedPassedCount := 2;
FSteps[9].ExpectedFailedCount := 0;
FSteps[9].CheckFinalization := TRUE;
FSteps[9].ExpectedFinalizationCount := 1;
FSteps[9].ExpectedCompletionCount := 1;
FSteps[9].ExpectedFinalResult := E_Result.Error;
FSteps[9].ExpectRuntimeHeld := TRUE;
FSteps[9].ExpectQuietCall := TRUE;
FSteps[9].ExpectedHookCount := 1;
FSteps[9].ExpectedHooks[1].Hook := E_LifecycleHook.Aggregate;
FSteps[9].ExpectedHooks[1].State := E_State.Completed;
FSteps[9].ExpectedHooks[1].Enabled := TRUE;
{endregion}

{region "10 - Reset clears the first result and competing requests"}
FSteps[10].ExpectedState := E_State.Idle;
FSteps[10].ExpectedResult := E_Result.NotEvaluated;
FSteps[10].ExpectedReady := TRUE;
FSteps[10].ExpectedPassedCount := 0;
FSteps[10].ExpectedFailedCount := 0;
FSteps[10].CheckFinalization := TRUE;
FSteps[10].ExpectedFinalizationCount := 1;
FSteps[10].ExpectedCompletionCount := 1;
FSteps[10].ExpectedFinalResult := E_Result.Error;
FSteps[10].RequestReset := TRUE;
FSteps[10].RequestStart := TRUE;
FSteps[10].RequestAbort := TRUE;
FSteps[10].ExpectRuntimeCleared := TRUE;
FSteps[10].ExpectedHookCount := 6;
FSteps[10].ExpectedHooks[1].Hook := E_LifecycleHook.Reset;
FSteps[10].ExpectedHooks[1].State := E_State.Reset;
FSteps[10].ExpectedHooks[1].Enabled := TRUE;
FSteps[10].ExpectedHooks[2].Hook := E_LifecycleHook.Abort;
FSteps[10].ExpectedHooks[2].State := E_State.Idle;
FSteps[10].ExpectedHooks[2].Enabled := FALSE;
FSteps[10].ExpectedHooks[3].Hook := E_LifecycleHook.Preparations;
FSteps[10].ExpectedHooks[3].State := E_State.Idle;
FSteps[10].ExpectedHooks[3].Enabled := FALSE;
FSteps[10].ExpectedHooks[4].Hook := E_LifecycleHook.Tests;
FSteps[10].ExpectedHooks[4].State := E_State.Idle;
FSteps[10].ExpectedHooks[4].Enabled := FALSE;
FSteps[10].ExpectedHooks[5].Hook := E_LifecycleHook.Assertions;
FSteps[10].ExpectedHooks[5].State := E_State.Idle;
FSteps[10].ExpectedHooks[5].Enabled := FALSE;
FSteps[10].ExpectedHooks[6].Hook := E_LifecycleHook.Aggregate;
FSteps[10].ExpectedHooks[6].State := E_State.Idle;
FSteps[10].ExpectedHooks[6].Enabled := TRUE;
{endregion}

{region "11 - Do not retain a Start from the Reset call"}
FSteps[11].ExpectedState := E_State.Idle;
FSteps[11].ExpectedResult := E_Result.NotEvaluated;
FSteps[11].ExpectedReady := TRUE;
FSteps[11].ExpectedPassedCount := 0;
FSteps[11].ExpectedFailedCount := 0;
FSteps[11].CheckFinalization := TRUE;
FSteps[11].ExpectedFinalizationCount := 1;
FSteps[11].ExpectedCompletionCount := 1;
FSteps[11].ExpectedFinalResult := E_Result.Error;
FSteps[11].ExpectRuntimeCleared := TRUE;
FSteps[11].ExpectQuietCall := TRUE;
FSteps[11].ExpectedHookCount := 5;
FSteps[11].ExpectedHooks[1].Hook := E_LifecycleHook.Abort;
FSteps[11].ExpectedHooks[1].State := E_State.Idle;
FSteps[11].ExpectedHooks[1].Enabled := FALSE;
FSteps[11].ExpectedHooks[2].Hook := E_LifecycleHook.Preparations;
FSteps[11].ExpectedHooks[2].State := E_State.Idle;
FSteps[11].ExpectedHooks[2].Enabled := FALSE;
FSteps[11].ExpectedHooks[3].Hook := E_LifecycleHook.Tests;
FSteps[11].ExpectedHooks[3].State := E_State.Idle;
FSteps[11].ExpectedHooks[3].Enabled := FALSE;
FSteps[11].ExpectedHooks[4].Hook := E_LifecycleHook.Assertions;
FSteps[11].ExpectedHooks[4].State := E_State.Idle;
FSteps[11].ExpectedHooks[4].Enabled := FALSE;
FSteps[11].ExpectedHooks[5].Hook := E_LifecycleHook.Aggregate;
FSteps[11].ExpectedHooks[5].State := E_State.Idle;
FSteps[11].ExpectedHooks[5].Enabled := TRUE;
{endregion}

{region "12 - Start a fresh second execution"}
FSteps[12].ExpectedState := E_State.Starting;
FSteps[12].ExpectedResult := E_Result.NotEvaluated;
FSteps[12].ExpectedReady := FALSE;
FSteps[12].ExpectedPassedCount := 0;
FSteps[12].ExpectedFailedCount := 0;
FSteps[12].CheckFinalization := TRUE;
FSteps[12].ExpectedFinalizationCount := 1;
FSteps[12].ExpectedCompletionCount := 1;
FSteps[12].ExpectedFinalResult := E_Result.Error;
FSteps[12].RequestStart := TRUE;
FSteps[12].ExpectedHookCount := 5;
FSteps[12].ExpectedHooks[1].Hook := E_LifecycleHook.Abort;
FSteps[12].ExpectedHooks[1].State := E_State.Starting;
FSteps[12].ExpectedHooks[1].Enabled := FALSE;
FSteps[12].ExpectedHooks[2].Hook := E_LifecycleHook.Preparations;
FSteps[12].ExpectedHooks[2].State := E_State.Starting;
FSteps[12].ExpectedHooks[2].Enabled := FALSE;
FSteps[12].ExpectedHooks[3].Hook := E_LifecycleHook.Tests;
FSteps[12].ExpectedHooks[3].State := E_State.Starting;
FSteps[12].ExpectedHooks[3].Enabled := FALSE;
FSteps[12].ExpectedHooks[4].Hook := E_LifecycleHook.Assertions;
FSteps[12].ExpectedHooks[4].State := E_State.Starting;
FSteps[12].ExpectedHooks[4].Enabled := FALSE;
FSteps[12].ExpectedHooks[5].Hook := E_LifecycleHook.Aggregate;
FSteps[12].ExpectedHooks[5].State := E_State.Starting;
FSteps[12].ExpectedHooks[5].Enabled := TRUE;
{endregion}

{region "13 - Both Assertions pass after Reset"}
FSteps[13].ExpectedState := E_State.Running;
FSteps[13].ExpectedResult := E_Result.NotEvaluated;
FSteps[13].ExpectedReady := FALSE;
FSteps[13].ExpectedPassedCount := 2;
FSteps[13].ExpectedFailedCount := 0;
FSteps[13].CheckFinalization := TRUE;
FSteps[13].ExpectedFinalizationCount := 1;
FSteps[13].ExpectedCompletionCount := 1;
FSteps[13].ExpectedFinalResult := E_Result.Error;
FSteps[13].ExpectedHookCount := 5;
FSteps[13].ExpectedHooks[1].Hook := E_LifecycleHook.Abort;
FSteps[13].ExpectedHooks[1].State := E_State.Running;
FSteps[13].ExpectedHooks[1].Enabled := FALSE;
FSteps[13].ExpectedHooks[2].Hook := E_LifecycleHook.Preparations;
FSteps[13].ExpectedHooks[2].State := E_State.Running;
FSteps[13].ExpectedHooks[2].Enabled := FALSE;
FSteps[13].ExpectedHooks[3].Hook := E_LifecycleHook.Tests;
FSteps[13].ExpectedHooks[3].State := E_State.Running;
FSteps[13].ExpectedHooks[3].Enabled := TRUE;
FSteps[13].ExpectedHooks[4].Hook := E_LifecycleHook.Assertions;
FSteps[13].ExpectedHooks[4].State := E_State.Running;
FSteps[13].ExpectedHooks[4].Enabled := TRUE;
FSteps[13].ExpectedHooks[5].Hook := E_LifecycleHook.Aggregate;
FSteps[13].ExpectedHooks[5].State := E_State.Running;
FSteps[13].ExpectedHooks[5].Enabled := TRUE;
{endregion}

{region "14 - Publish a new successful finalization"}
FSteps[14].ExpectedState := E_State.Completing;
FSteps[14].ExpectedResult := E_Result.Passed;
FSteps[14].ExpectedReady := FALSE;
FSteps[14].ExpectedPassedCount := 2;
FSteps[14].ExpectedFailedCount := 0;
FSteps[14].FinishTests := TRUE;
FSteps[14].CheckFinalization := TRUE;
FSteps[14].ExpectedFinalizationCount := 2;
FSteps[14].ExpectedCompletionCount := 1;
FSteps[14].ExpectedFinalResult := E_Result.Passed;
FSteps[14].ExpectedHookCount := 5;
FSteps[14].ExpectedHooks[1].Hook := E_LifecycleHook.Abort;
FSteps[14].ExpectedHooks[1].State := E_State.Running;
FSteps[14].ExpectedHooks[1].Enabled := FALSE;
FSteps[14].ExpectedHooks[2].Hook := E_LifecycleHook.Preparations;
FSteps[14].ExpectedHooks[2].State := E_State.Running;
FSteps[14].ExpectedHooks[2].Enabled := FALSE;
FSteps[14].ExpectedHooks[3].Hook := E_LifecycleHook.Tests;
FSteps[14].ExpectedHooks[3].State := E_State.Running;
FSteps[14].ExpectedHooks[3].Enabled := TRUE;
FSteps[14].ExpectedHooks[4].Hook := E_LifecycleHook.Assertions;
FSteps[14].ExpectedHooks[4].State := E_State.Completing;
FSteps[14].ExpectedHooks[4].Enabled := FALSE;
FSteps[14].ExpectedHooks[5].Hook := E_LifecycleHook.Aggregate;
FSteps[14].ExpectedHooks[5].State := E_State.Completing;
FSteps[14].ExpectedHooks[5].Enabled := TRUE;
{endregion}

{region "15 - Complete the second execution"}
FSteps[15].ExpectedState := E_State.Completed;
FSteps[15].ExpectedResult := E_Result.Passed;
FSteps[15].ExpectedReady := FALSE;
FSteps[15].ExpectedPassedCount := 2;
FSteps[15].ExpectedFailedCount := 0;
FSteps[15].ExpectRuntimeHeld := TRUE;
FSteps[15].CheckFinalization := TRUE;
FSteps[15].ExpectedFinalizationCount := 2;
FSteps[15].ExpectedCompletionCount := 2;
FSteps[15].ExpectedFinalResult := E_Result.Passed;
FSteps[15].ExpectedHookCount := 1;
FSteps[15].ExpectedHooks[1].Hook := E_LifecycleHook.Aggregate;
FSteps[15].ExpectedHooks[1].State := E_State.Completed;
FSteps[15].ExpectedHooks[1].Enabled := TRUE;
{endregion}

{region "16 - Do not repeat second-run finalization"}
FSteps[16].ExpectedState := E_State.Completed;
FSteps[16].ExpectedResult := E_Result.Passed;
FSteps[16].ExpectedReady := FALSE;
FSteps[16].ExpectedPassedCount := 2;
FSteps[16].ExpectedFailedCount := 0;
FSteps[16].ExpectQuietCall := TRUE;
FSteps[16].ExpectRuntimeHeld := TRUE;
FSteps[16].CheckFinalization := TRUE;
FSteps[16].ExpectedFinalizationCount := 2;
FSteps[16].ExpectedCompletionCount := 2;
FSteps[16].ExpectedFinalResult := E_Result.Passed;
FSteps[16].ExpectedHookCount := 1;
FSteps[16].ExpectedHooks[1].Hook := E_LifecycleHook.Aggregate;
FSteps[16].ExpectedHooks[1].State := E_State.Completed;
FSteps[16].ExpectedHooks[1].Enabled := TRUE;
{endregion}
END_METHOD

END_FUNCTION_BLOCK

// ---- SelfTests/TestCases/TestSuite_TestCaseLifecycle/Test_LifecycleRepeatAfterAbort.TcPOU
{region 'Documentation'}
(*!
<summary>Checks stable Abort completion, one-shot finalization and a fresh successful run after Reset.</summary>
*)
{endregion}
FUNCTION_BLOCK Test_LifecycleRepeatAfterAbort EXTENDS TestCaseLifecycleTestBase

SUPER^();

{region 'Documentation'}
(*!
<summary>Defines two independent run outcomes and cumulative event expectations across Reset.</summary>
*)
{endregion}
METHOD PROTECTED ConfigureScenario
FSubjectPreparationCount := 0;
FSubjectTestCount := 1;
FStepCount := 15;

{region "01 - Reset establishes the initial Idle state"}
FSteps[1].ExpectedState := E_State.Idle;
FSteps[1].ExpectedResult := E_Result.NotEvaluated;
FSteps[1].ExpectedReady := TRUE;
FSteps[1].ExpectedPassedCount := 0;
FSteps[1].ExpectedFailedCount := 0;
FSteps[1].RequestReset := TRUE;
FSteps[1].ExpectRuntimeCleared := TRUE;
FSteps[1].CheckFinalization := TRUE;
FSteps[1].ExpectedFinalizationCount := 0;
FSteps[1].ExpectedCompletionCount := 0;
FSteps[1].ExpectedFinalResult := E_Result.Abort;
FSteps[1].ExpectedHookCount := 6;
FSteps[1].ExpectedHooks[1].Hook := E_LifecycleHook.Reset;
FSteps[1].ExpectedHooks[1].State := E_State.Reset;
FSteps[1].ExpectedHooks[1].Enabled := TRUE;
FSteps[1].ExpectedHooks[2].Hook := E_LifecycleHook.Abort;
FSteps[1].ExpectedHooks[2].State := E_State.Idle;
FSteps[1].ExpectedHooks[2].Enabled := FALSE;
FSteps[1].ExpectedHooks[3].Hook := E_LifecycleHook.Preparations;
FSteps[1].ExpectedHooks[3].State := E_State.Idle;
FSteps[1].ExpectedHooks[3].Enabled := FALSE;
FSteps[1].ExpectedHooks[4].Hook := E_LifecycleHook.Tests;
FSteps[1].ExpectedHooks[4].State := E_State.Idle;
FSteps[1].ExpectedHooks[4].Enabled := FALSE;
FSteps[1].ExpectedHooks[5].Hook := E_LifecycleHook.Assertions;
FSteps[1].ExpectedHooks[5].State := E_State.Idle;
FSteps[1].ExpectedHooks[5].Enabled := FALSE;
FSteps[1].ExpectedHooks[6].Hook := E_LifecycleHook.Aggregate;
FSteps[1].ExpectedHooks[6].State := E_State.Idle;
FSteps[1].ExpectedHooks[6].Enabled := TRUE;
{endregion}

{region "02 - Start the first execution"}
FSteps[2].ExpectedState := E_State.Starting;
FSteps[2].ExpectedResult := E_Result.NotEvaluated;
FSteps[2].ExpectedReady := FALSE;
FSteps[2].ExpectedPassedCount := 0;
FSteps[2].ExpectedFailedCount := 0;
FSteps[2].RequestStart := TRUE;
FSteps[2].CheckFinalization := TRUE;
FSteps[2].ExpectedFinalizationCount := 0;
FSteps[2].ExpectedCompletionCount := 0;
FSteps[2].ExpectedFinalResult := E_Result.Abort;
FSteps[2].ExpectedHookCount := 5;
FSteps[2].ExpectedHooks[1].Hook := E_LifecycleHook.Abort;
FSteps[2].ExpectedHooks[1].State := E_State.Starting;
FSteps[2].ExpectedHooks[1].Enabled := FALSE;
FSteps[2].ExpectedHooks[2].Hook := E_LifecycleHook.Preparations;
FSteps[2].ExpectedHooks[2].State := E_State.Starting;
FSteps[2].ExpectedHooks[2].Enabled := FALSE;
FSteps[2].ExpectedHooks[3].Hook := E_LifecycleHook.Tests;
FSteps[2].ExpectedHooks[3].State := E_State.Starting;
FSteps[2].ExpectedHooks[3].Enabled := FALSE;
FSteps[2].ExpectedHooks[4].Hook := E_LifecycleHook.Assertions;
FSteps[2].ExpectedHooks[4].State := E_State.Starting;
FSteps[2].ExpectedHooks[4].Enabled := FALSE;
FSteps[2].ExpectedHooks[5].Hook := E_LifecycleHook.Aggregate;
FSteps[2].ExpectedHooks[5].State := E_State.Starting;
FSteps[2].ExpectedHooks[5].Enabled := TRUE;
{endregion}

{region "03 - Evaluate both child Assertions"}
FSteps[3].ExpectedState := E_State.Running;
FSteps[3].ExpectedResult := E_Result.NotEvaluated;
FSteps[3].ExpectedReady := FALSE;
FSteps[3].ExpectedPassedCount := 2;
FSteps[3].ExpectedFailedCount := 0;
FSteps[3].AssertionCondition := TRUE;
FSteps[3].CheckFinalization := TRUE;
FSteps[3].ExpectedFinalizationCount := 0;
FSteps[3].ExpectedCompletionCount := 0;
FSteps[3].ExpectedFinalResult := E_Result.Abort;
FSteps[3].ExpectedHookCount := 5;
FSteps[3].ExpectedHooks[1].Hook := E_LifecycleHook.Abort;
FSteps[3].ExpectedHooks[1].State := E_State.Running;
FSteps[3].ExpectedHooks[1].Enabled := FALSE;
FSteps[3].ExpectedHooks[2].Hook := E_LifecycleHook.Preparations;
FSteps[3].ExpectedHooks[2].State := E_State.Running;
FSteps[3].ExpectedHooks[2].Enabled := FALSE;
FSteps[3].ExpectedHooks[3].Hook := E_LifecycleHook.Tests;
FSteps[3].ExpectedHooks[3].State := E_State.Running;
FSteps[3].ExpectedHooks[3].Enabled := TRUE;
FSteps[3].ExpectedHooks[4].Hook := E_LifecycleHook.Assertions;
FSteps[3].ExpectedHooks[4].State := E_State.Running;
FSteps[3].ExpectedHooks[4].Enabled := TRUE;
FSteps[3].ExpectedHooks[5].Hook := E_LifecycleHook.Aggregate;
FSteps[3].ExpectedHooks[5].State := E_State.Running;
FSteps[3].ExpectedHooks[5].Enabled := TRUE;
{endregion}

{region "04 - Acknowledge explicit Abort"}
FSteps[4].ExpectedState := E_State.Completing;
FSteps[4].ExpectedResult := E_Result.Abort;
FSteps[4].ExpectedReady := FALSE;
FSteps[4].ExpectedPassedCount := 2;
FSteps[4].ExpectedFailedCount := 0;
FSteps[4].RequestAbort := TRUE;
FSteps[4].CheckFinalization := TRUE;
FSteps[4].ExpectedFinalizationCount := 1;
FSteps[4].ExpectedCompletionCount := 0;
FSteps[4].ExpectedFinalResult := E_Result.Abort;
FSteps[4].ExpectedHookCount := 5;
FSteps[4].ExpectedHooks[1].Hook := E_LifecycleHook.Abort;
FSteps[4].ExpectedHooks[1].State := E_State.Aborting;
FSteps[4].ExpectedHooks[1].Enabled := TRUE;
FSteps[4].ExpectedHooks[2].Hook := E_LifecycleHook.Preparations;
FSteps[4].ExpectedHooks[2].State := E_State.Completing;
FSteps[4].ExpectedHooks[2].Enabled := FALSE;
FSteps[4].ExpectedHooks[3].Hook := E_LifecycleHook.Tests;
FSteps[4].ExpectedHooks[3].State := E_State.Completing;
FSteps[4].ExpectedHooks[3].Enabled := FALSE;
FSteps[4].ExpectedHooks[4].Hook := E_LifecycleHook.Assertions;
FSteps[4].ExpectedHooks[4].State := E_State.Completing;
FSteps[4].ExpectedHooks[4].Enabled := FALSE;
FSteps[4].ExpectedHooks[5].Hook := E_LifecycleHook.Aggregate;
FSteps[4].ExpectedHooks[5].State := E_State.Completing;
FSteps[4].ExpectedHooks[5].Enabled := TRUE;
{endregion}

{region "05 - Observe the final Completed transition"}
FSteps[5].ExpectedState := E_State.Completed;
FSteps[5].ExpectedResult := E_Result.Abort;
FSteps[5].ExpectedReady := FALSE;
FSteps[5].ExpectedPassedCount := 2;
FSteps[5].ExpectedFailedCount := 0;
FSteps[5].CheckFinalization := TRUE;
FSteps[5].ExpectedFinalizationCount := 1;
FSteps[5].ExpectedCompletionCount := 1;
FSteps[5].ExpectedFinalResult := E_Result.Abort;
FSteps[5].ExpectRuntimeHeld := TRUE;
FSteps[5].ExpectedHookCount := 1;
FSteps[5].ExpectedHooks[1].Hook := E_LifecycleHook.Aggregate;
FSteps[5].ExpectedHooks[1].State := E_State.Completed;
FSteps[5].ExpectedHooks[1].Enabled := TRUE;
{endregion}

{region "06 - Ignore processing inputs while Completed"}
FSteps[6].ExpectedState := E_State.Completed;
FSteps[6].ExpectedResult := E_Result.Abort;
FSteps[6].ExpectedReady := FALSE;
FSteps[6].ExpectedPassedCount := 2;
FSteps[6].ExpectedFailedCount := 0;
FSteps[6].CheckFinalization := TRUE;
FSteps[6].ExpectedFinalizationCount := 1;
FSteps[6].ExpectedCompletionCount := 1;
FSteps[6].ExpectedFinalResult := E_Result.Abort;
FSteps[6].ExpectRuntimeHeld := TRUE;
FSteps[6].ExpectQuietCall := TRUE;
FSteps[6].Ready := FALSE;
FSteps[6].ResetError := TRUE;
FSteps[6].AbortError := TRUE;
FSteps[6].TestError := TRUE;
FSteps[6].PreparationError := TRUE;
FSteps[6].AdvancePreparation := TRUE;
FSteps[6].FinishPreparations := TRUE;
FSteps[6].AdvanceTest := TRUE;
FSteps[6].FinishTests := TRUE;
FSteps[6].AssertionCondition := FALSE;
FSteps[6].ExpectedHookCount := 1;
FSteps[6].ExpectedHooks[1].Hook := E_LifecycleHook.Aggregate;
FSteps[6].ExpectedHooks[1].State := E_State.Completed;
FSteps[6].ExpectedHooks[1].Enabled := TRUE;
{endregion}

{region "07 - Consume Start and Abort without restarting"}
FSteps[7].ExpectedState := E_State.Completed;
FSteps[7].ExpectedResult := E_Result.Abort;
FSteps[7].ExpectedReady := FALSE;
FSteps[7].ExpectedPassedCount := 2;
FSteps[7].ExpectedFailedCount := 0;
FSteps[7].CheckFinalization := TRUE;
FSteps[7].ExpectedFinalizationCount := 1;
FSteps[7].ExpectedCompletionCount := 1;
FSteps[7].ExpectedFinalResult := E_Result.Abort;
FSteps[7].ExpectRuntimeHeld := TRUE;
FSteps[7].RequestStart := TRUE;
FSteps[7].RequestAbort := TRUE;
FSteps[7].ExpectedHookCount := 1;
FSteps[7].ExpectedHooks[1].Hook := E_LifecycleHook.Aggregate;
FSteps[7].ExpectedHooks[1].State := E_State.Completed;
FSteps[7].ExpectedHooks[1].Enabled := TRUE;
{endregion}

{region "08 - Remain quiet after rejected terminal requests"}
FSteps[8].ExpectedState := E_State.Completed;
FSteps[8].ExpectedResult := E_Result.Abort;
FSteps[8].ExpectedReady := FALSE;
FSteps[8].ExpectedPassedCount := 2;
FSteps[8].ExpectedFailedCount := 0;
FSteps[8].CheckFinalization := TRUE;
FSteps[8].ExpectedFinalizationCount := 1;
FSteps[8].ExpectedCompletionCount := 1;
FSteps[8].ExpectedFinalResult := E_Result.Abort;
FSteps[8].ExpectRuntimeHeld := TRUE;
FSteps[8].ExpectQuietCall := TRUE;
FSteps[8].ExpectedHookCount := 1;
FSteps[8].ExpectedHooks[1].Hook := E_LifecycleHook.Aggregate;
FSteps[8].ExpectedHooks[1].State := E_State.Completed;
FSteps[8].ExpectedHooks[1].Enabled := TRUE;
{endregion}

{region "09 - Reset clears the first result and competing requests"}
FSteps[9].ExpectedState := E_State.Idle;
FSteps[9].ExpectedResult := E_Result.NotEvaluated;
FSteps[9].ExpectedReady := TRUE;
FSteps[9].ExpectedPassedCount := 0;
FSteps[9].ExpectedFailedCount := 0;
FSteps[9].CheckFinalization := TRUE;
FSteps[9].ExpectedFinalizationCount := 1;
FSteps[9].ExpectedCompletionCount := 1;
FSteps[9].ExpectedFinalResult := E_Result.Abort;
FSteps[9].RequestReset := TRUE;
FSteps[9].RequestStart := TRUE;
FSteps[9].RequestAbort := TRUE;
FSteps[9].ExpectRuntimeCleared := TRUE;
FSteps[9].ExpectedHookCount := 6;
FSteps[9].ExpectedHooks[1].Hook := E_LifecycleHook.Reset;
FSteps[9].ExpectedHooks[1].State := E_State.Reset;
FSteps[9].ExpectedHooks[1].Enabled := TRUE;
FSteps[9].ExpectedHooks[2].Hook := E_LifecycleHook.Abort;
FSteps[9].ExpectedHooks[2].State := E_State.Idle;
FSteps[9].ExpectedHooks[2].Enabled := FALSE;
FSteps[9].ExpectedHooks[3].Hook := E_LifecycleHook.Preparations;
FSteps[9].ExpectedHooks[3].State := E_State.Idle;
FSteps[9].ExpectedHooks[3].Enabled := FALSE;
FSteps[9].ExpectedHooks[4].Hook := E_LifecycleHook.Tests;
FSteps[9].ExpectedHooks[4].State := E_State.Idle;
FSteps[9].ExpectedHooks[4].Enabled := FALSE;
FSteps[9].ExpectedHooks[5].Hook := E_LifecycleHook.Assertions;
FSteps[9].ExpectedHooks[5].State := E_State.Idle;
FSteps[9].ExpectedHooks[5].Enabled := FALSE;
FSteps[9].ExpectedHooks[6].Hook := E_LifecycleHook.Aggregate;
FSteps[9].ExpectedHooks[6].State := E_State.Idle;
FSteps[9].ExpectedHooks[6].Enabled := TRUE;
{endregion}

{region "10 - Do not retain a Start from the Reset call"}
FSteps[10].ExpectedState := E_State.Idle;
FSteps[10].ExpectedResult := E_Result.NotEvaluated;
FSteps[10].ExpectedReady := TRUE;
FSteps[10].ExpectedPassedCount := 0;
FSteps[10].ExpectedFailedCount := 0;
FSteps[10].CheckFinalization := TRUE;
FSteps[10].ExpectedFinalizationCount := 1;
FSteps[10].ExpectedCompletionCount := 1;
FSteps[10].ExpectedFinalResult := E_Result.Abort;
FSteps[10].ExpectRuntimeCleared := TRUE;
FSteps[10].ExpectQuietCall := TRUE;
FSteps[10].ExpectedHookCount := 5;
FSteps[10].ExpectedHooks[1].Hook := E_LifecycleHook.Abort;
FSteps[10].ExpectedHooks[1].State := E_State.Idle;
FSteps[10].ExpectedHooks[1].Enabled := FALSE;
FSteps[10].ExpectedHooks[2].Hook := E_LifecycleHook.Preparations;
FSteps[10].ExpectedHooks[2].State := E_State.Idle;
FSteps[10].ExpectedHooks[2].Enabled := FALSE;
FSteps[10].ExpectedHooks[3].Hook := E_LifecycleHook.Tests;
FSteps[10].ExpectedHooks[3].State := E_State.Idle;
FSteps[10].ExpectedHooks[3].Enabled := FALSE;
FSteps[10].ExpectedHooks[4].Hook := E_LifecycleHook.Assertions;
FSteps[10].ExpectedHooks[4].State := E_State.Idle;
FSteps[10].ExpectedHooks[4].Enabled := FALSE;
FSteps[10].ExpectedHooks[5].Hook := E_LifecycleHook.Aggregate;
FSteps[10].ExpectedHooks[5].State := E_State.Idle;
FSteps[10].ExpectedHooks[5].Enabled := TRUE;
{endregion}

{region "11 - Start a fresh second execution"}
FSteps[11].ExpectedState := E_State.Starting;
FSteps[11].ExpectedResult := E_Result.NotEvaluated;
FSteps[11].ExpectedReady := FALSE;
FSteps[11].ExpectedPassedCount := 0;
FSteps[11].ExpectedFailedCount := 0;
FSteps[11].CheckFinalization := TRUE;
FSteps[11].ExpectedFinalizationCount := 1;
FSteps[11].ExpectedCompletionCount := 1;
FSteps[11].ExpectedFinalResult := E_Result.Abort;
FSteps[11].RequestStart := TRUE;
FSteps[11].ExpectedHookCount := 5;
FSteps[11].ExpectedHooks[1].Hook := E_LifecycleHook.Abort;
FSteps[11].ExpectedHooks[1].State := E_State.Starting;
FSteps[11].ExpectedHooks[1].Enabled := FALSE;
FSteps[11].ExpectedHooks[2].Hook := E_LifecycleHook.Preparations;
FSteps[11].ExpectedHooks[2].State := E_State.Starting;
FSteps[11].ExpectedHooks[2].Enabled := FALSE;
FSteps[11].ExpectedHooks[3].Hook := E_LifecycleHook.Tests;
FSteps[11].ExpectedHooks[3].State := E_State.Starting;
FSteps[11].ExpectedHooks[3].Enabled := FALSE;
FSteps[11].ExpectedHooks[4].Hook := E_LifecycleHook.Assertions;
FSteps[11].ExpectedHooks[4].State := E_State.Starting;
FSteps[11].ExpectedHooks[4].Enabled := FALSE;
FSteps[11].ExpectedHooks[5].Hook := E_LifecycleHook.Aggregate;
FSteps[11].ExpectedHooks[5].State := E_State.Starting;
FSteps[11].ExpectedHooks[5].Enabled := TRUE;
{endregion}

{region "12 - Both Assertions pass after Reset"}
FSteps[12].ExpectedState := E_State.Running;
FSteps[12].ExpectedResult := E_Result.NotEvaluated;
FSteps[12].ExpectedReady := FALSE;
FSteps[12].ExpectedPassedCount := 2;
FSteps[12].ExpectedFailedCount := 0;
FSteps[12].CheckFinalization := TRUE;
FSteps[12].ExpectedFinalizationCount := 1;
FSteps[12].ExpectedCompletionCount := 1;
FSteps[12].ExpectedFinalResult := E_Result.Abort;
FSteps[12].ExpectedHookCount := 5;
FSteps[12].ExpectedHooks[1].Hook := E_LifecycleHook.Abort;
FSteps[12].ExpectedHooks[1].State := E_State.Running;
FSteps[12].ExpectedHooks[1].Enabled := FALSE;
FSteps[12].ExpectedHooks[2].Hook := E_LifecycleHook.Preparations;
FSteps[12].ExpectedHooks[2].State := E_State.Running;
FSteps[12].ExpectedHooks[2].Enabled := FALSE;
FSteps[12].ExpectedHooks[3].Hook := E_LifecycleHook.Tests;
FSteps[12].ExpectedHooks[3].State := E_State.Running;
FSteps[12].ExpectedHooks[3].Enabled := TRUE;
FSteps[12].ExpectedHooks[4].Hook := E_LifecycleHook.Assertions;
FSteps[12].ExpectedHooks[4].State := E_State.Running;
FSteps[12].ExpectedHooks[4].Enabled := TRUE;
FSteps[12].ExpectedHooks[5].Hook := E_LifecycleHook.Aggregate;
FSteps[12].ExpectedHooks[5].State := E_State.Running;
FSteps[12].ExpectedHooks[5].Enabled := TRUE;
{endregion}

{region "13 - Publish a new successful finalization"}
FSteps[13].ExpectedState := E_State.Completing;
FSteps[13].ExpectedResult := E_Result.Passed;
FSteps[13].ExpectedReady := FALSE;
FSteps[13].ExpectedPassedCount := 2;
FSteps[13].ExpectedFailedCount := 0;
FSteps[13].FinishTests := TRUE;
FSteps[13].CheckFinalization := TRUE;
FSteps[13].ExpectedFinalizationCount := 2;
FSteps[13].ExpectedCompletionCount := 1;
FSteps[13].ExpectedFinalResult := E_Result.Passed;
FSteps[13].ExpectedHookCount := 5;
FSteps[13].ExpectedHooks[1].Hook := E_LifecycleHook.Abort;
FSteps[13].ExpectedHooks[1].State := E_State.Running;
FSteps[13].ExpectedHooks[1].Enabled := FALSE;
FSteps[13].ExpectedHooks[2].Hook := E_LifecycleHook.Preparations;
FSteps[13].ExpectedHooks[2].State := E_State.Running;
FSteps[13].ExpectedHooks[2].Enabled := FALSE;
FSteps[13].ExpectedHooks[3].Hook := E_LifecycleHook.Tests;
FSteps[13].ExpectedHooks[3].State := E_State.Running;
FSteps[13].ExpectedHooks[3].Enabled := TRUE;
FSteps[13].ExpectedHooks[4].Hook := E_LifecycleHook.Assertions;
FSteps[13].ExpectedHooks[4].State := E_State.Completing;
FSteps[13].ExpectedHooks[4].Enabled := FALSE;
FSteps[13].ExpectedHooks[5].Hook := E_LifecycleHook.Aggregate;
FSteps[13].ExpectedHooks[5].State := E_State.Completing;
FSteps[13].ExpectedHooks[5].Enabled := TRUE;
{endregion}

{region "14 - Complete the second execution"}
FSteps[14].ExpectedState := E_State.Completed;
FSteps[14].ExpectedResult := E_Result.Passed;
FSteps[14].ExpectedReady := FALSE;
FSteps[14].ExpectedPassedCount := 2;
FSteps[14].ExpectedFailedCount := 0;
FSteps[14].ExpectRuntimeHeld := TRUE;
FSteps[14].CheckFinalization := TRUE;
FSteps[14].ExpectedFinalizationCount := 2;
FSteps[14].ExpectedCompletionCount := 2;
FSteps[14].ExpectedFinalResult := E_Result.Passed;
FSteps[14].ExpectedHookCount := 1;
FSteps[14].ExpectedHooks[1].Hook := E_LifecycleHook.Aggregate;
FSteps[14].ExpectedHooks[1].State := E_State.Completed;
FSteps[14].ExpectedHooks[1].Enabled := TRUE;
{endregion}

{region "15 - Do not repeat second-run finalization"}
FSteps[15].ExpectedState := E_State.Completed;
FSteps[15].ExpectedResult := E_Result.Passed;
FSteps[15].ExpectedReady := FALSE;
FSteps[15].ExpectedPassedCount := 2;
FSteps[15].ExpectedFailedCount := 0;
FSteps[15].ExpectQuietCall := TRUE;
FSteps[15].ExpectRuntimeHeld := TRUE;
FSteps[15].CheckFinalization := TRUE;
FSteps[15].ExpectedFinalizationCount := 2;
FSteps[15].ExpectedCompletionCount := 2;
FSteps[15].ExpectedFinalResult := E_Result.Passed;
FSteps[15].ExpectedHookCount := 1;
FSteps[15].ExpectedHooks[1].Hook := E_LifecycleHook.Aggregate;
FSteps[15].ExpectedHooks[1].State := E_State.Completed;
FSteps[15].ExpectedHooks[1].Enabled := TRUE;
{endregion}
END_METHOD

END_FUNCTION_BLOCK

// ---- SelfTests/TestSuites/TestSuite_Orchestrator.TcPOU
{region 'Documentation'}
(*!
<summary>Verifies common Orchestrator behavior through isolated subjects with a Serial arrangement.</summary>
*)
{endregion}
FUNCTION_BLOCK TestSuite_Orchestrator EXTENDS TestSuiteBase
VAR
    FShiftedBounds : Test_OrchestratorShiftedBounds;
    FNegativeBounds : Test_OrchestratorNegativeBounds;
    FUnusedCapacity : Test_OrchestratorUnusedCapacity;
    FSingleChild : Test_OrchestratorSingleChild;
    FIdleReadiness : Test_OrchestratorIdleReadiness;
    FMissingStartReaction : Test_OrchestratorMissingStartReaction;
    FChildError : Test_OrchestratorChildError;
    FUnexpectedAbort : Test_OrchestratorUnexpectedAbort;
    FAbortInterruption : Test_OrchestratorAbortInterruption;
    FIdleInterruption : Test_OrchestratorIdleInterruption;
    FResetInterruption : Test_OrchestratorResetInterruption;
    FResetContinuesAfterError : Test_OrchestratorResetContinuesAfterError;
    FRepeatAfterReset : Test_OrchestratorRepeatAfterReset;
    FExecutionCapacityWait : Test_OrchestratorExecutionCapacityWait;
    FResetCapacityWait : Test_OrchestratorResetCapacityWait;
    FExecutionBudgetError : Test_OrchestratorExecutionBudgetError;
    FTestCases : ARRAY[1..TestCaseCapacity] OF I_TestCase;
END_VAR
VAR CONSTANT
    TestCaseCapacity : UINT := 16;
END_VAR

SUPER^();

{region 'Documentation'}
(*!
<summary>Initializes and registers the owned orchestration scenarios in deterministic order.</summary>
*)
{endregion}
METHOD PROTECTED Configure
VAR_IN_OUT
    // SA0167: Borrowed builder; VAR_IN_OUT creates no temporary instance.
    {attribute 'analysis' := '-167'}
    Builder : TestSuiteConfigurationBuilder; //! Borrowed owner configuration builder used only during this Configure call; register this owner's concrete children.
END_VAR
VAR
    TestConfig : ST_TestCaseConfig;
END_VAR
Builder.Initialize(Mode := E_OrchestrationMode.Serial,
    TestCases := FTestCases);

FShiftedBounds.Initialize(Parent := THIS^,
    TestName := 'ShiftedBounds',
    Config := TestConfig);
Builder.Register(TestCase := FShiftedBounds);

FNegativeBounds.Initialize(Parent := THIS^,
    TestName := 'NegativeBounds',
    Config := TestConfig);
Builder.Register(TestCase := FNegativeBounds);

FUnusedCapacity.Initialize(Parent := THIS^,
    TestName := 'UnusedCapacity',
    Config := TestConfig);
Builder.Register(TestCase := FUnusedCapacity);

FSingleChild.Initialize(Parent := THIS^,
    TestName := 'SingleChild',
    Config := TestConfig);
Builder.Register(TestCase := FSingleChild);

FIdleReadiness.Initialize(Parent := THIS^,
    TestName := 'IdleReadiness',
    Config := TestConfig);
Builder.Register(TestCase := FIdleReadiness);

FMissingStartReaction.Initialize(Parent := THIS^,
    TestName := 'MissingStartReaction',
    Config := TestConfig);
Builder.Register(TestCase := FMissingStartReaction);

FChildError.Initialize(Parent := THIS^,
    TestName := 'ChildError',
    Config := TestConfig);
Builder.Register(TestCase := FChildError);

FUnexpectedAbort.Initialize(Parent := THIS^,
    TestName := 'UnexpectedAbort',
    Config := TestConfig);
Builder.Register(TestCase := FUnexpectedAbort);

FAbortInterruption.Initialize(Parent := THIS^,
    TestName := 'AbortInterruption',
    Config := TestConfig);
Builder.Register(TestCase := FAbortInterruption);

FIdleInterruption.Initialize(Parent := THIS^,
    TestName := 'IdleInterruption',
    Config := TestConfig);
Builder.Register(TestCase := FIdleInterruption);

FResetInterruption.Initialize(Parent := THIS^,
    TestName := 'ResetInterruption',
    Config := TestConfig);
Builder.Register(TestCase := FResetInterruption);

FResetContinuesAfterError.Initialize(Parent := THIS^,
    TestName := 'ResetContinuesAfterError',
    Config := TestConfig);
Builder.Register(TestCase := FResetContinuesAfterError);

FRepeatAfterReset.Initialize(Parent := THIS^,
    TestName := 'RepeatAfterReset',
    Config := TestConfig);
Builder.Register(TestCase := FRepeatAfterReset);

FExecutionCapacityWait.Initialize(Parent := THIS^,
    TestName := 'ExecutionCapacityWait',
    Config := TestConfig);
Builder.Register(TestCase := FExecutionCapacityWait);

FResetCapacityWait.Initialize(Parent := THIS^,
    TestName := 'ResetCapacityWait',
    Config := TestConfig);
Builder.Register(TestCase := FResetCapacityWait);

FExecutionBudgetError.Initialize(Parent := THIS^,
    TestName := 'ExecutionBudgetError',
    Config := TestConfig);
Builder.Register(TestCase := FExecutionBudgetError);
END_METHOD

{region 'Documentation'}
(*!
<summary>Returns the registered Test Case from the same array used during configuration.</summary>
*)
{endregion}
METHOD PUBLIC GetTestCase : I_TestCase //! Typed child interface at the original array index; zero when no entry is available.
VAR_INPUT
    Index : DINT; //! Original occupied child-array index, rather than an ordinal position.
END_VAR
GetTestCase := 0;
IF (ChildCount = 0) OR (Index < ChildArrayLowerBound)
    OR (DINT_TO_LINT(Index) >= DINT_TO_LINT(ChildArrayLowerBound) + UINT_TO_LINT(ChildCount)) THEN
    RETURN;
END_IF;

GetTestCase := FTestCases[Index];
END_METHOD

{region 'Documentation'}
(*!
<summary>Calls each owned Test Case once per initialized Suite cycle, including completion.</summary>
*)
{endregion}
METHOD PROTECTED ProcessTestCases
FShiftedBounds();
FNegativeBounds();
FUnusedCapacity();
FSingleChild();
FIdleReadiness();
FMissingStartReaction();
FChildError();
FUnexpectedAbort();
FAbortInterruption();
FIdleInterruption();
FResetInterruption();
FResetContinuesAfterError();
FRepeatAfterReset();
FExecutionCapacityWait();
FResetCapacityWait();
FExecutionBudgetError();
END_METHOD

END_FUNCTION_BLOCK

// ---- SelfTests/TestCases/TestSuite_Orchestrator/Test_OrchestratorShiftedBounds.TcPOU
{region 'Documentation'}
(*!
<summary>Checks the same execution trace with actual indices 7 through 9.</summary>
*)
{endregion}
FUNCTION_BLOCK Test_OrchestratorShiftedBounds EXTENDS OrchestrationTestBase

SUPER^();

{region 'Documentation'}
(*!
<summary>Defines this scenario independently of the subject's internal fields.</summary>
*)
{endregion}
METHOD PROTECTED ConfigureScenario
FArrayLayout := E_OrchestrationArrayLayout.Shifted;
FChildCount := 3;
ConfigureStandardSequence();
END_METHOD

END_FUNCTION_BLOCK

// ---- SelfTests/Helper/Orchestration/OrchestrationTestBase.TcPOU
{region 'Documentation'}
(*!
<summary>Runs explicit per-cycle scenarios against the real shared Orchestrator.</summary>
<description>

Roles

FSubject is the unchanged production Orchestrator with local diagnostic capture.
FChildren are interface doubles, not TestCaseBase copies. FCollection exposes the
registered prefix at the selected array's real indices; unused capacity stays empty.
Only the outer Assertions publish into the normal selftest Event Stream.

Scenario composition

ConfigureScenario assigns FChildSlots before fixture initialization. Defaults are
1, 2, 3 for Serial; Parallel scenarios assign slot 1 to every participating child.
Each row states MaxActiveChildCount, defaulting to the existing Serial limit of one.
Activity includes this call's Start request and prior active child observations.
The limit applies during Execution; per-child request checks still allow only one Start.

One checkpoint per task cycle

ConfigureScenario supplies independent child observations and helper expectations.
ProcessTests clears call evidence and installs reservation responses for the current row,
calls the helper once, then each registered child once.
Accepted responses are the default. Unaccepted reservation expectations count additional
WaitingForCapacity or Error attempts without Start/Reset; they do not imply dispatch.
Child requests are recorded before the script's next observation is applied.
ProcessAssertions compares this cycle before the next checkpoint can advance.
No extra call is made to acknowledge a Start; the next helper call sees the prior child call.

Trace and scope

FTrace retains before/after observations, requests, releases and helper outputs.
The table is an explicit regression trace for this call order, not a second scheduler.
Reservation markers check interface ordering, not real Event Buffer budget arithmetic.
Outer Reset rebuilds the isolated fixture. The ordinary subject Reset is a separate task.

Errors and interruptions

ExpectedDiagnosticCount is cumulative within the scenario, including across subject Reset.
Held errors must not generate repeated events. Captured payloads are checked by
classification and owner context, not by diagnostic message wording.
Reset/Abort requests and task-specific completion are explicit per-cycle expectations;
Reset completion and helper readiness remain distinct observations.
</description>
*)
{endregion}
FUNCTION_BLOCK ABSTRACT OrchestrationTestBase EXTENDS TestCaseBase
VAR
    FSubject : OrchestratorProbe;
    FCollection : OrchestrationCollectionDouble;
    FChildren : ARRAY[1..3] OF OrchestrationChildDouble;
    FOrdinaryChildren : ARRAY[1..3] OF I_Orchestratable;
    FShiftedChildren : ARRAY[7..9] OF I_Orchestratable;
    FNegativeChildren : ARRAY[-3..-1] OF I_Orchestratable;
    FSpareChildren : ARRAY[1..6] OF I_Orchestratable;
    FArrayLayout : E_OrchestrationArrayLayout := E_OrchestrationArrayLayout.Ordinary;
    FChildCount : UINT := 3;
    FChildSlots : ARRAY[1..3] OF UINT := [1, 2, 3];
    FSteps : ARRAY[1..StepCapacity] OF ST_OrchestrationStep;
    FTrace : ARRAY[1..StepCapacity] OF ST_OrchestrationCycle;
    FStepCount : INT;
    FStepIndex : INT := 1;
    FCheckPerformed : BOOL;
    FObservationReady : BOOL;
    FFixtureValid : BOOL;
    FCapture : EventBuffer;
    FEvents : ARRAY[1..CaptureLength] OF ST_Event;
    FCaptureFifo : ST_FifoStatus;
    FCaptureStatus : ST_EventBufferStatus;
    FCheckRequests : AssertTrue;
    FCheckOtherRequests : AssertTrue;
    FCheckReservations : AssertTrue;
    FCheckChildCalls : AssertTrue;
    FCheckCollectionAccess : AssertTrue;
    FCheckActiveChildren : AssertTrue;
    FCheckSlot : AssertEqual_UInt;
    FCheckCompletion : AssertEqual_Bool;
    FCheckReady : AssertEqual_Bool;
    FCheckTask : AssertEqual_Int;
    FCheckResult : AssertEqual_Int;
    FCheckDiagnostics : AssertEqual_UDInt;
    FCheckTaskStatus : AssertTrue;
    FCheckDiagnosticPayload : AssertTrue;
END_VAR
VAR CONSTANT
    StepCapacity : INT := 24;
    CaptureLength : UINT := 32;
END_VAR

SUPER^();

{region 'Documentation'}
(*!
<summary>Contributes every outer Assertion once without running the isolated scheduler.</summary>
*)
{endregion}
METHOD PROTECTED AggregateResults
VAR_INPUT
    Aggregator : I_ResultAggregator; //! Borrowed result sink owned by the outer Test Case; add this test's checking Assertions without resetting or retaining the sink.
END_VAR
Aggregator.AddProvider(Provider := FCheckRequests);
Aggregator.AddProvider(Provider := FCheckOtherRequests);
Aggregator.AddProvider(Provider := FCheckReservations);
Aggregator.AddProvider(Provider := FCheckChildCalls);
Aggregator.AddProvider(Provider := FCheckCollectionAccess);
Aggregator.AddProvider(Provider := FCheckActiveChildren);
Aggregator.AddProvider(Provider := FCheckSlot);
Aggregator.AddProvider(Provider := FCheckCompletion);
Aggregator.AddProvider(Provider := FCheckReady);
Aggregator.AddProvider(Provider := FCheckTask);
Aggregator.AddProvider(Provider := FCheckResult);
Aggregator.AddProvider(Provider := FCheckDiagnostics);
Aggregator.AddProvider(Provider := FCheckTaskStatus);
Aggregator.AddProvider(Provider := FCheckDiagnosticPayload);
END_METHOD

{region 'Documentation'}
(*!
<summary>Validates isolated Framework diagnostics without depending on their message wording.</summary>
<description>
The local buffer is neither deleted nor overwritten during a scenario.
Sequence count detects missing or repeated publication. This check validates
classification, owner context and storage integrity of every captured entry.
</description>
*)
{endregion}
METHOD PRIVATE AreDiagnosticsValid : BOOL //! TRUE when capture accounting and every retained diagnostic match the expected Framework error context.
VAR
    Index : UINT;
    Diagnostic : REFERENCE TO ST_Event;
    ExpectedName : STRING(GVL_Constants.NameLength);
END_VAR
AreDiagnosticsValid := FALSE;
IF FCaptureFifo.ConfigError OR FCaptureFifo.IndexError
    OR (FCaptureStatus.LostEventCount <> 0)
    OR (FCaptureFifo.ElementCount >= CaptureLength)
    OR (FCaptureFifo.IndexOut <> 1)
    OR (FCaptureStatus.SequenceId <> UINT_TO_UDINT(FCaptureFifo.ElementCount)) THEN
    RETURN;
END_IF;

ExpectedName := CONCAT(Name, '.Orchestrator');
FOR Index := 1 TO FCaptureFifo.ElementCount DO
    Diagnostic REF= FEvents[Index];
    IF (Diagnostic.SequenceId <> UINT_TO_UDINT(Index))
        OR (Diagnostic.OwnerScope <> E_OwnerScope.Framework)
        OR (Diagnostic.EventType <> E_EventType.Framework)
        OR (Diagnostic.Severity <> E_EventSeverity.Error)
        OR (Diagnostic.State <> E_State.Error)
        OR (Diagnostic.Result <> E_Result.NotEvaluated)
        OR (Diagnostic.Name <> ExpectedName)
        OR (Diagnostic.ResourceName <> '')
        OR (Diagnostic.Message = '') THEN
        RETURN;
    END_IF;
END_FOR;
AreDiagnosticsValid := TRUE;
END_METHOD

{region 'Documentation'}
(*!
<summary>Includes scenario bounds, fixture binding and evaluating Assertions in initialization validity.</summary>
*)
{endregion}
METHOD PROTECTED CheckInitialization : BOOL //! TRUE when the inherited initialization check and this concrete fixture check both accept the setup.
CheckInitialization := FALSE;
IF NOT SUPER^.CheckInitialization() THEN
    RETURN;
END_IF;
IF NOT FFixtureValid OR (FStepCount < 1) OR (FStepCount > StepCapacity) THEN
    RETURN;
END_IF;
IF NOT FCheckRequests.IsInitialized
    OR NOT FCheckOtherRequests.IsInitialized
    OR NOT FCheckReservations.IsInitialized
    OR NOT FCheckChildCalls.IsInitialized
    OR NOT FCheckCollectionAccess.IsInitialized
    OR NOT FCheckActiveChildren.IsInitialized
    OR NOT FCheckSlot.IsInitialized
    OR NOT FCheckCompletion.IsInitialized
    OR NOT FCheckReady.IsInitialized
    OR NOT FCheckTask.IsInitialized
    OR NOT FCheckResult.IsInitialized
    OR NOT FCheckDiagnostics.IsInitialized
    OR NOT FCheckTaskStatus.IsInitialized
    OR NOT FCheckDiagnosticPayload.IsInitialized THEN
    RETURN;
END_IF;
CheckInitialization := TRUE;
END_METHOD

{region 'Documentation'}
(*!
<summary>Defines scenario tables and initializes the isolated fixture and outer Assertions.</summary>
*)
{endregion}
METHOD PROTECTED Configure
VAR
    Index : INT;
    EmptyStep : ST_OrchestrationStep;
END_VAR
FOR Index := 1 TO StepCapacity DO
    FSteps[Index] := EmptyStep;
END_FOR;
FStepCount := 0;
FChildCount := 3;
FArrayLayout := E_OrchestrationArrayLayout.Ordinary;
FOR Index := 1 TO 3 DO
    FChildSlots[Index] := INT_TO_UINT(Index);
END_FOR;
ConfigureScenario();
FPreparationStateCount := 0;
FTestStateCount := FStepCount;
FFixtureValid := InitializeFixture();
FCheckRequests.Initialize(Parent := THIS^,
    AssertionName := 'Requests');
FCheckOtherRequests.Initialize(Parent := THIS^,
    AssertionName := 'OtherRequests');
FCheckReservations.Initialize(Parent := THIS^,
    AssertionName := 'Reservations');
FCheckChildCalls.Initialize(Parent := THIS^,
    AssertionName := 'ChildCalls');
FCheckCollectionAccess.Initialize(Parent := THIS^,
    AssertionName := 'CollectionAccess');
FCheckActiveChildren.Initialize(Parent := THIS^,
    AssertionName := 'ActiveChildren');
FCheckSlot.Initialize(Parent := THIS^,
    AssertionName := 'Slot');
FCheckCompletion.Initialize(Parent := THIS^,
    AssertionName := 'Completion');
FCheckReady.Initialize(Parent := THIS^,
    AssertionName := 'Ready');
FCheckTask.Initialize(Parent := THIS^,
    AssertionName := 'Task');
FCheckResult.Initialize(Parent := THIS^,
    AssertionName := 'Result');
FCheckDiagnostics.Initialize(Parent := THIS^,
    AssertionName := 'Diagnostics');
FCheckTaskStatus.Initialize(Parent := THIS^,
    AssertionName := 'TaskStatus');
FCheckDiagnosticPayload.Initialize(Parent := THIS^,
    AssertionName := 'DiagnosticPayload');
END_METHOD

{region 'Documentation'}
(*!
<summary>Defines collection layout, child slots, population and independent cyclic expectations.</summary>
*)
{endregion}
METHOD PROTECTED ABSTRACT ConfigureScenario
END_METHOD

{region 'Documentation'}
(*!
<summary>Defines the same A-B-C request trace for collection-index and capacity variants.</summary>
*)
{endregion}
METHOD PROTECTED ConfigureStandardSequence
FStepCount := 12;

{region "Cycle 01 - Idle readiness"}
FSteps[1].Task := E_OrchestratorTask.Idle;
FSteps[1].ExpectedReady := TRUE;
{endregion}

{region "Cycle 02 - Start child 1"}
FSteps[2].Children[1].State := E_State.Running;
FSteps[2].Children[1].Ready := FALSE;
FSteps[2].ExpectedStartChild := 1;
FSteps[2].ExpectedSlot := 1;
FSteps[2].ExpectedReservations[1] := 1;
{endregion}

{region "Cycle 03 - Child progress"}
FSteps[3].Children[1].State := E_State.Running;
FSteps[3].Children[1].Ready := FALSE;
FSteps[3].ExpectedSlot := 1;
FSteps[3].ExpectedReservations[1] := 1;
{endregion}

{region "Cycle 04 - Child progress"}
FSteps[4].Children[1].State := E_State.Completed;
FSteps[4].Children[1].Ready := FALSE;
FSteps[4].Children[1].Complete := TRUE;
FSteps[4].Children[1].Result := E_Result.Passed;
FSteps[4].ExpectedSlot := 1;
FSteps[4].ExpectedReservations[1] := 1;
{endregion}

{region "Cycle 05 - Reconcile completed child 1"}
FSteps[5].Children[1].State := E_State.Completed;
FSteps[5].Children[1].Ready := FALSE;
FSteps[5].Children[1].Complete := TRUE;
FSteps[5].Children[1].Result := E_Result.Passed;
FSteps[5].ExpectedSlot := 2;
FSteps[5].ExpectedReleasedEntries[1] := 1;
{endregion}

{region "Cycle 06 - Start child 2"}
FSteps[6].Children[1].State := E_State.Completed;
FSteps[6].Children[1].Ready := FALSE;
FSteps[6].Children[1].Complete := TRUE;
FSteps[6].Children[1].Result := E_Result.Passed;
FSteps[6].Children[2].State := E_State.Running;
FSteps[6].Children[2].Ready := FALSE;
FSteps[6].ExpectedStartChild := 2;
FSteps[6].ExpectedSlot := 2;
FSteps[6].ExpectedReservations[2] := 1;
{endregion}

{region "Cycle 07 - Child progress"}
FSteps[7].Children[1].State := E_State.Completed;
FSteps[7].Children[1].Ready := FALSE;
FSteps[7].Children[1].Complete := TRUE;
FSteps[7].Children[1].Result := E_Result.Passed;
FSteps[7].Children[2].State := E_State.Completed;
FSteps[7].Children[2].Ready := FALSE;
FSteps[7].Children[2].Complete := TRUE;
FSteps[7].Children[2].Result := E_Result.Passed;
FSteps[7].ExpectedSlot := 2;
FSteps[7].ExpectedReservations[2] := 1;
{endregion}

{region "Cycle 08 - Reconcile completed child 2"}
FSteps[8].Children[1].State := E_State.Completed;
FSteps[8].Children[1].Ready := FALSE;
FSteps[8].Children[1].Complete := TRUE;
FSteps[8].Children[1].Result := E_Result.Passed;
FSteps[8].Children[2].State := E_State.Completed;
FSteps[8].Children[2].Ready := FALSE;
FSteps[8].Children[2].Complete := TRUE;
FSteps[8].Children[2].Result := E_Result.Passed;
FSteps[8].ExpectedSlot := 3;
FSteps[8].ExpectedReleasedEntries[2] := 1;
{endregion}

{region "Cycle 09 - Start child 3"}
FSteps[9].Children[1].State := E_State.Completed;
FSteps[9].Children[1].Ready := FALSE;
FSteps[9].Children[1].Complete := TRUE;
FSteps[9].Children[1].Result := E_Result.Passed;
FSteps[9].Children[2].State := E_State.Completed;
FSteps[9].Children[2].Ready := FALSE;
FSteps[9].Children[2].Complete := TRUE;
FSteps[9].Children[2].Result := E_Result.Passed;
FSteps[9].Children[3].State := E_State.Running;
FSteps[9].Children[3].Ready := FALSE;
FSteps[9].ExpectedStartChild := 3;
FSteps[9].ExpectedSlot := 3;
FSteps[9].ExpectedReservations[3] := 1;
{endregion}

{region "Cycle 10 - Child progress"}
FSteps[10].Children[1].State := E_State.Completed;
FSteps[10].Children[1].Ready := FALSE;
FSteps[10].Children[1].Complete := TRUE;
FSteps[10].Children[1].Result := E_Result.Passed;
FSteps[10].Children[2].State := E_State.Completed;
FSteps[10].Children[2].Ready := FALSE;
FSteps[10].Children[2].Complete := TRUE;
FSteps[10].Children[2].Result := E_Result.Passed;
FSteps[10].Children[3].State := E_State.Completed;
FSteps[10].Children[3].Ready := FALSE;
FSteps[10].Children[3].Complete := TRUE;
FSteps[10].Children[3].Result := E_Result.Passed;
FSteps[10].ExpectedSlot := 3;
FSteps[10].ExpectedReservations[3] := 1;
{endregion}

{region "Cycle 11 - Completed observation"}
FSteps[11].Children[1].State := E_State.Completed;
FSteps[11].Children[1].Ready := FALSE;
FSteps[11].Children[1].Complete := TRUE;
FSteps[11].Children[1].Result := E_Result.Passed;
FSteps[11].Children[2].State := E_State.Completed;
FSteps[11].Children[2].Ready := FALSE;
FSteps[11].Children[2].Complete := TRUE;
FSteps[11].Children[2].Result := E_Result.Passed;
FSteps[11].Children[3].State := E_State.Completed;
FSteps[11].Children[3].Ready := FALSE;
FSteps[11].Children[3].Complete := TRUE;
FSteps[11].Children[3].Result := E_Result.Passed;
FSteps[11].ExpectedReleasedEntries[3] := 1;
FSteps[11].ExpectedFinished := TRUE;
{endregion}

{region "Cycle 12 - Completed observation"}
FSteps[12].Children[1].State := E_State.Completed;
FSteps[12].Children[1].Ready := FALSE;
FSteps[12].Children[1].Complete := TRUE;
FSteps[12].Children[1].Result := E_Result.Passed;
FSteps[12].Children[2].State := E_State.Completed;
FSteps[12].Children[2].Ready := FALSE;
FSteps[12].Children[2].Complete := TRUE;
FSteps[12].Children[2].Result := E_Result.Passed;
FSteps[12].Children[3].State := E_State.Completed;
FSteps[12].Children[3].Ready := FALSE;
FSteps[12].Children[3].Complete := TRUE;
FSteps[12].Children[3].Result := E_Result.Passed;
FSteps[12].ExpectedFinished := TRUE;
{endregion}
END_METHOD

{region 'Documentation'}
(*!
<summary>Rebuilds local capture, children, collection and helper before any scenario call.</summary>
*)
{endregion}
METHOD PRIVATE InitializeFixture : BOOL //! TRUE when local capture, array layout, collection and real helper initialization all succeed.
VAR
    Position : UINT;
    Index : INT;
    EmptyCycle : ST_OrchestrationCycle;
    CollectionValid : BOOL;
END_VAR
InitializeFixture := FALSE;
FStepIndex := 1;
FCheckPerformed := FALSE;
FObservationReady := FALSE;
FOR Index := 1 TO StepCapacity DO
    FTrace[Index] := EmptyCycle;
END_FOR;
IF (FChildCount < 1) OR (FChildCount > 3) THEN
    RETURN;
END_IF;
IF NOT FCapture.Initialize(Buffer := FEvents,
    FifoControl := FCaptureFifo,
    Status := FCaptureStatus) THEN
    RETURN;
END_IF;

FOR Position := 1 TO 3 DO
    FChildren[Position].Initialize(Name := CONCAT('Child', UINT_TO_STRING(Position)),
        Slot := FChildSlots[Position]);
    FOrdinaryChildren[Position] := 0;
    FShiftedChildren[UINT_TO_INT(Position) + 6] := 0;
    FNegativeChildren[UINT_TO_INT(Position) - 4] := 0;
END_FOR;
FOR Position := 1 TO 6 DO
    FSpareChildren[Position] := 0;
END_FOR;
FOR Position := 1 TO FChildCount DO
    CASE FArrayLayout OF
        E_OrchestrationArrayLayout.Ordinary:
            FOrdinaryChildren[Position] := FChildren[Position];
        E_OrchestrationArrayLayout.Shifted:
            FShiftedChildren[UINT_TO_INT(Position) + 6] := FChildren[Position];
        E_OrchestrationArrayLayout.Negative:
            FNegativeChildren[UINT_TO_INT(Position) - 4] := FChildren[Position];
        E_OrchestrationArrayLayout.SpareCapacity:
            FSpareChildren[Position] := FChildren[Position];
    ELSE
        RETURN;
    END_CASE;
END_FOR;
CASE FArrayLayout OF
    E_OrchestrationArrayLayout.Ordinary:
        CollectionValid := FCollection.Initialize(Count := FChildCount,
            Children := FOrdinaryChildren);
    E_OrchestrationArrayLayout.Shifted:
        CollectionValid := FCollection.Initialize(Count := FChildCount,
            Children := FShiftedChildren);
    E_OrchestrationArrayLayout.Negative:
        CollectionValid := FCollection.Initialize(Count := FChildCount,
            Children := FNegativeChildren);
    E_OrchestrationArrayLayout.SpareCapacity:
        CollectionValid := FCollection.Initialize(Count := FChildCount,
            Children := FSpareChildren);
ELSE
    RETURN;
END_CASE;
IF NOT CollectionValid THEN
    RETURN;
END_IF;

FSubject.BindPublisher(Publisher := FCapture);
InitializeFixture := FSubject.Initialize(Collection := FCollection,
    Name := Name);
END_METHOD

{region 'Documentation'}
(*!
<summary>Completes outer Abort; isolated children have no external resource effects.</summary>
*)
{endregion}
METHOD PROTECTED ProcessAbort
VAR_INPUT
    Enable : BOOL; //! Phase permission supplied by the owning Test Case; FALSE does not authorize progression, while observation may continue.
END_VAR
IF Enable THEN
    CompleteAbort();
END_IF;
END_METHOD

{region 'Documentation'}
(*!
<summary>Checks each explicit row; latched Assertion results retain any earlier mismatch.</summary>
*)
{endregion}
METHOD PROTECTED ProcessAssertions
VAR_INPUT
    Enable : BOOL; //! Phase permission supplied by the owning Test Case; FALSE does not authorize progression, while observation may continue.
END_VAR
VAR
    EvaluateChecks : BOOL;
    Position : UINT;
    ExpectedStarts : UINT;
    ExpectedResets : UINT;
    RequestsMatch : BOOL;
    OtherRequestsMatch : BOOL;
    ReservationsMatch : BOOL;
    ChildCallsMatch : BOOL;
END_VAR
EvaluateChecks := Enable AND FObservationReady;
RequestsMatch := TRUE;
OtherRequestsMatch := TRUE;
ReservationsMatch := FTrace[FStepIndex].RequestsDidNotChangeState;
ChildCallsMatch := FTrace[FStepIndex].HelperDidNotCallChildren;
FOR Position := 1 TO FChildCount DO
    ExpectedStarts := BOOL_TO_UINT(FSteps[FStepIndex].ExpectedStartChild = Position);
    ExpectedResets := BOOL_TO_UINT(FSteps[FStepIndex].ExpectedResetChild = Position);
    RequestsMatch := RequestsMatch
        AND (FTrace[FStepIndex].Calls[Position].StartCount = ExpectedStarts);
    OtherRequestsMatch := OtherRequestsMatch
        AND (FTrace[FStepIndex].Calls[Position].ResetCount = ExpectedResets)
        AND (FTrace[FStepIndex].Calls[Position].AbortCount = FSteps[FStepIndex].ExpectedAbortRequests[Position])
        AND (FTrace[FStepIndex].Calls[Position].ResetReservationCount = ExpectedResets
            + FSteps[FStepIndex].ExpectedUnacceptedResetReservations[Position]);
    ReservationsMatch := ReservationsMatch
        AND (FTrace[FStepIndex].Calls[Position].ExecutionReservationCount = ExpectedStarts
            + FSteps[FStepIndex].ExpectedUnacceptedExecutionReservations[Position])
        AND NOT FTrace[FStepIndex].Calls[Position].StartWithoutReservation
        AND NOT FTrace[FStepIndex].Calls[Position].ResetWithoutReservation
        AND (FTrace[FStepIndex].Reservations[Position] = FSteps[FStepIndex].ExpectedReservations[Position])
        AND (FTrace[FStepIndex].Calls[Position].ReleasedEntryCount = FSteps[FStepIndex].ExpectedReleasedEntries[Position]);
    ChildCallsMatch := ChildCallsMatch AND (FTrace[FStepIndex].Calls[Position].BodyCount = 1);
END_FOR;

FCheckRequests(Enable := EvaluateChecks,
    State := State,
    IN := RequestsMatch);
FCheckOtherRequests(Enable := EvaluateChecks,
    State := State,
    IN := OtherRequestsMatch);
FCheckReservations(Enable := EvaluateChecks,
    State := State,
    IN := ReservationsMatch);
FCheckChildCalls(Enable := EvaluateChecks,
    State := State,
    IN := ChildCallsMatch);
FCheckCollectionAccess(Enable := EvaluateChecks,
    State := State,
    IN := NOT FCollection.InvalidAccess AND NOT FCollection.TraceOverflow
        AND (FCollection.ReadCount > 0));
FCheckActiveChildren(Enable := EvaluateChecks,
    State := State,
    IN := (FSteps[FStepIndex].Task <> E_OrchestratorTask.Execution)
        OR (FTrace[FStepIndex].ActiveChildCount <= FSteps[FStepIndex].MaxActiveChildCount));
FCheckSlot(Enable := EvaluateChecks,
    State := State,
    IN := FTrace[FStepIndex].ActiveSlot,
    Expected := FSteps[FStepIndex].ExpectedSlot);
FCheckCompletion(Enable := EvaluateChecks,
    State := State,
    IN := FTrace[FStepIndex].ExecutionFinished,
    Expected := FSteps[FStepIndex].ExpectedFinished);
FCheckReady(Enable := EvaluateChecks,
    State := State,
    IN := FTrace[FStepIndex].Ready,
    Expected := FSteps[FStepIndex].ExpectedReady);
FCheckTask(Enable := EvaluateChecks,
    State := State,
    IN := TO_INT(FTrace[FStepIndex].Task),
    Expected := TO_INT(FSteps[FStepIndex].Task));
FCheckResult(Enable := EvaluateChecks,
    State := State,
    IN := TO_INT(FTrace[FStepIndex].Result),
    Expected := TO_INT(FSteps[FStepIndex].ExpectedResult));
FCheckDiagnostics(Enable := EvaluateChecks,
    State := State,
    IN := FCaptureStatus.SequenceId,
    Expected := FSteps[FStepIndex].ExpectedDiagnosticCount);
FCheckTaskStatus(Enable := EvaluateChecks,
    State := State,
    IN := (FTrace[FStepIndex].ResetFinished = FSteps[FStepIndex].ExpectedResetFinished)
        AND (FTrace[FStepIndex].AbortFinished = FSteps[FStepIndex].ExpectedAbortFinished)
        AND (FTrace[FStepIndex].TaskComplete = (FSteps[FStepIndex].ExpectedFinished
            OR FSteps[FStepIndex].ExpectedResetFinished OR FSteps[FStepIndex].ExpectedAbortFinished))
        AND (FTrace[FStepIndex].ResetActive = (FSteps[FStepIndex].Task = E_OrchestratorTask.Reset))
        AND (FTrace[FStepIndex].ExecutionActive = (FSteps[FStepIndex].Task = E_OrchestratorTask.Execution))
        AND (FTrace[FStepIndex].AbortActive = (FSteps[FStepIndex].Task = E_OrchestratorTask.Abort)));
FCheckDiagnosticPayload(Enable := EvaluateChecks,
    State := State,
    IN := AreDiagnosticsValid());

IF EvaluateChecks
    AND FCheckRequests.EvaluationActive
    AND FCheckOtherRequests.EvaluationActive
    AND FCheckReservations.EvaluationActive
    AND FCheckChildCalls.EvaluationActive
    AND FCheckCollectionAccess.EvaluationActive
    AND FCheckActiveChildren.EvaluationActive
    AND FCheckSlot.EvaluationActive
    AND FCheckCompletion.EvaluationActive
    AND FCheckReady.EvaluationActive
    AND FCheckTask.EvaluationActive
    AND FCheckResult.EvaluationActive
    AND FCheckDiagnostics.EvaluationActive
    AND FCheckTaskStatus.EvaluationActive
    AND FCheckDiagnosticPayload.EvaluationActive THEN
    FCheckPerformed := TRUE;
END_IF;
END_METHOD

{region 'Documentation'}
(*!
<summary>No outer Preparation is required; child views are local scenario data.</summary>
*)
{endregion}
METHOD PROTECTED ProcessPreparations
VAR_INPUT
    // SA0033: Required hook with no Preparation work.
    {attribute 'analysis' := '-33'}
    Enable : BOOL; //! Phase permission supplied by the owning Test Case; FALSE does not authorize progression, while observation may continue.
END_VAR
END_METHOD

{region 'Documentation'}
(*!
<summary>Clears outer checks and rebuilds the fixture; does not simulate a subject Reset task.</summary>
*)
{endregion}
METHOD PROTECTED ProcessReset
FCheckRequests.Reset();
FCheckOtherRequests.Reset();
FCheckReservations.Reset();
FCheckChildCalls.Reset();
FCheckCollectionAccess.Reset();
FCheckActiveChildren.Reset();
FCheckSlot.Reset();
FCheckCompletion.Reset();
FCheckReady.Reset();
FCheckTask.Reset();
FCheckResult.Reset();
FCheckDiagnostics.Reset();
FCheckTaskStatus.Reset();
FCheckDiagnosticPayload.Reset();
FFixtureValid := InitializeFixture();
IF NOT FFixtureValid THEN
    Error(Message := 'Orchestration fixture setup failed.');
END_IF;
CompleteReset();
END_METHOD

{region 'Documentation'}
(*!
<summary>Runs the helper before children exactly once per checkpoint and retains evidence.</summary>
*)
{endregion}
METHOD PROTECTED ProcessTests
VAR_INPUT
    Enable : BOOL; //! Phase permission supplied by the owning Test Case; FALSE does not authorize progression, while observation may continue.
END_VAR
VAR
    Position : UINT;
    BeforeHelper : ARRAY[1..3] OF ST_OrchestrationObservation;
    AfterHelper : ST_OrchestrationObservation;
    Calls : ST_OrchestrationCalls;
END_VAR
FObservationReady := FALSE;
IF NOT Enable THEN
    RETURN;
END_IF;

IF FCheckPerformed THEN
    FCheckPerformed := FALSE;
    IF FStepIndex = FStepCount THEN
        CompleteTests();
        RETURN;
    END_IF;
    FStepIndex := FStepIndex + 1;
    NextTestState();
    IF NOT IsTestingActive THEN
        RETURN;
    END_IF;
END_IF;

FOR Position := 1 TO FChildCount DO
    FChildren[Position].BeginCycle(ExecutionReservationResult := FSteps[FStepIndex].ExecutionReservationResults[Position],
        ResetReservationResult := FSteps[FStepIndex].ResetReservationResults[Position]);
    BeforeHelper[Position] := FChildren[Position].Observation;
END_FOR;

FSubject(Task := FSteps[FStepIndex].Task);
FTrace[FStepIndex].ActiveSlot := FSubject.ActiveSlot;
FTrace[FStepIndex].ExecutionFinished := FSubject.IsExecutionFinished;
FTrace[FStepIndex].ResetFinished := FSubject.IsResetFinished;
FTrace[FStepIndex].AbortFinished := FSubject.IsAbortFinished;
FTrace[FStepIndex].TaskComplete := FSubject.IsComplete;
FTrace[FStepIndex].ResetActive := FSubject.IsResetActive;
FTrace[FStepIndex].ExecutionActive := FSubject.IsExecutionActive;
FTrace[FStepIndex].AbortActive := FSubject.IsAbortActive;
FTrace[FStepIndex].Ready := FSubject.IsReady;
FTrace[FStepIndex].Result := FSubject.Result;
FTrace[FStepIndex].Task := FSubject.CurrentTask;
FTrace[FStepIndex].HelperDidNotCallChildren := TRUE;
FTrace[FStepIndex].RequestsDidNotChangeState := TRUE;

// Inspect the helper boundary before applying any new child observation.
FOR Position := 1 TO FChildCount DO
    Calls := FChildren[Position].Calls;
    FTrace[FStepIndex].HelperDidNotCallChildren :=
        FTrace[FStepIndex].HelperDidNotCallChildren AND (Calls.BodyCount = 0);
    AfterHelper := FChildren[Position].Observation;
    FTrace[FStepIndex].BeforeChildren[Position] := AfterHelper;
    FTrace[FStepIndex].RequestsDidNotChangeState :=
        FTrace[FStepIndex].RequestsDidNotChangeState
        AND (AfterHelper.State = BeforeHelper[Position].State)
        AND (AfterHelper.Result = BeforeHelper[Position].Result)
        AND (AfterHelper.Ready = BeforeHelper[Position].Ready)
        AND (AfterHelper.Complete = BeforeHelper[Position].Complete);
    FTrace[FStepIndex].Reservations[Position] := FChildren[Position].ReservedEntryCount;
    IF (Calls.StartCount > 0)
        OR ((AfterHelper.State >= E_State.Starting) AND (AfterHelper.State <= E_State.Completing)) THEN
        FTrace[FStepIndex].ActiveChildCount := FTrace[FStepIndex].ActiveChildCount + 1;
    END_IF;
END_FOR;

FOR Position := 1 TO FChildCount DO
    FChildren[Position](ObservationInput := FSteps[FStepIndex].Children[Position]);
    FTrace[FStepIndex].Calls[Position] := FChildren[Position].Calls;
    FTrace[FStepIndex].AfterChildren[Position] := FChildren[Position].Observation;
END_FOR;
FObservationReady := TRUE;
END_METHOD

END_FUNCTION_BLOCK

// ---- SelfTests/Helper/Orchestration/OrchestratorProbe.TcPOU
{region 'Documentation'}
(*!
<summary>Uses the real scheduling algorithm with a pre-use local publisher binding.</summary>
*)
{endregion}
FUNCTION_BLOCK OrchestratorProbe EXTENDS Orchestrator

SUPER^(Task := Task);

{region 'Documentation'}
(*!
<summary>Binds isolated diagnostics before Initialize or any cyclic use.</summary>
*)
{endregion}
METHOD PUBLIC BindPublisher
VAR_INPUT
    Publisher : I_EventPublisher; //! Nonzero isolated event publisher retained before subject initialization; keep it alive through all subject use.
END_VAR
FEventPublisher := Publisher;
END_METHOD

END_FUNCTION_BLOCK

// ---- SelfTests/Helper/Orchestration/OrchestrationCollectionDouble.TcPOU
{region 'Documentation'}
(*!
<summary>Copies a small fixed child view and records actual-index access by the helper.</summary>
<description>
Initialize reads real bounds from the fixture's selected fixed array and copies only
its registered prefix. The copy is intentional test-double storage, not a production
registry or retained array pointer. GetChild translates the original index without
calling a child. Invalid access and trace overflow remain observable.
</description>
*)
{endregion}
FUNCTION_BLOCK OrchestrationCollectionDouble IMPLEMENTS I_OrchestratableCollection
VAR
    FChildren : ARRAY[1..ChildCapacity] OF I_Orchestratable;
    FLowerBound : DINT;
    FUpperBound : DINT;
    FCount : UINT;
    FReadIndices : ARRAY[1..ReadCapacity] OF DINT;
    FReadCount : UINT;
    FInvalidAccess : BOOL;
    FTraceOverflow : BOOL;
END_VAR
VAR CONSTANT
    ChildCapacity : UINT := 3;
    ReadCapacity : UINT := 512;
END_VAR

{region 'Documentation'}
(*!
<summary>Actual input-array lower bound.</summary>
*)
{endregion}
{attribute 'monitoring' := 'call'}
PROPERTY PUBLIC ChildArrayLowerBound : DINT //! Actual input-array lower bound.
GET
ChildArrayLowerBound := FLowerBound;
END_GET
END_PROPERTY

{region 'Documentation'}
(*!
<summary>Actual input-array capacity upper bound.</summary>
*)
{endregion}
{attribute 'monitoring' := 'call'}
PROPERTY PUBLIC ChildArrayUpperBound : DINT //! Actual input-array capacity upper bound.
GET
ChildArrayUpperBound := FUpperBound;
END_GET
END_PROPERTY

